(* IEC 61131-3 sources: daoli-st-library/DL_Motion (part 22) *)

(* ---- FB_DL_ElectronicCam.st ---- *)
(*==============================================================================
 * 组件名称 (Component)  : FB_DL_ElectronicCam
 * 所属子库 (Sublibrary) : DL_Motion
 * 当前版本 (Version)    : 1.0.0
 * 组件分类 (Category)   : 功能块（FUNCTION_BLOCK）· 多轴同步耦合族 · 电子凸轮
 * 兼容性   (Platform)   : CODESYS 3.5 / TwinCAT 3 / 汇川 InoProShop / Schneider
 *                         Machine Expert；仅依赖 Standard.library
 *                         （R_TRIG / LIMIT / MIN / MAX / ABS / 类型转换），零厂商方言
 * 接口依赖 (Depends)    : I_DL_MotionAxis / E_DL_AxisState（既有契约，Round 05，零修改）
 * 功能描述 (Function)   : 电子凸轮（PLCopen 凸轮耦合语义的 clean-room 独立实现）。
 *                         以「主轴相位归一化 → 分段线性表插值 → 缩放与偏移」四段
 *                         链计算从轴目标位置，支持周期 / 非周期两种运行方式、主
 *                         轴相位固定偏移与运行相位微调（飞剪切点补偿）、表单调性
 *                         校验与啮合过渡。
 * 设计要点 (Key notes)  :
 *   ① 相位归一化用「截断取整 + 条件加减」实现小数部分，绝不对负数取模，
 *      保证负向主轴时相位仍落在 0.0..1.0。
 *   ② 表查找为线性扫描 + 防死锁计数器；插值斜率计算前强制判分母，重合点保底
 *      取左值（重合已在啮合前由单调性校验拦截）。
 *   ③ 啮合前对全表做一次性扫描（点数 / 单调性 / 非有限值），运行中只校验当前
 *      区间，避免每拍全表扫描拖长任务周期。
 *   ④ 对轴接口每拍至多一次方法调用：定位指令与减速指令在同一拍互斥。
 * 开源溯源 (Origin)     : 原创实现，clean-room。语义来源为汇川 / CODESYS SoftMotion
 *                         公开指令手册的凸轮耦合页面、ABB AC500 PLCopen 库公开
 *                         帮助页、PLC 技术网公开实战帖与非周期追剪技术文
 *                         （来源编号 RAW_NOTES S-2）。
 *                         「借鉴对象的许可说明」：上述对象全部为公开发布但受版权
 *                         保护的帮助文档 / 论坛教程 / 技术文章，属「可免费查阅、
 *                         仅借鉴语义」类别；本实现未复制任何厂商源码、未使用其
 *                         凸轮表 XML 格式，引脚命名、表结构、插值实现、单调性
 *                         校验、故障码与状态机 100% 自有设计。
 * 验收向量 (Acceptance) :
 *   V1 三点表（0/0、180/90、360/0）周期运行：从轴位置连续，无阶跃跳变；
 *   V2 非周期走完表尾 → eComplete 且 bEndOfProfile 置位，等新啮合沿重启；
 *   V3 主轴点等值（非单调）→ 啮合沿受理时锁存 0004_0261；
 *   V4 nCamPoints = 1 → 锁存 0004_0260；
 *   V5 反向主轴 + bDirNegative = TRUE 正常同步；bDirNegative = FALSE 时停留
 *      eWaiting 并出信息级 0004_0140；
 *   V6 fPhaseShift 步进 5 mm → 切点前移且出信息级 0004_0142；
 *   V7 缩放填 0 → 回默认 1.0 并出信息级 0004_0141；
 *   V8 表值含非有限值 → 锁存 0004_0263；
 *   V9 运行中途插入跟踪脉冲 bTrack：重采样相位基准、退回 eIdle（公约 0.1）。
 * 已知限制 (Limits)     :
 *   ① 从轴定位经轴接口每拍一次下发，同步精度受扫描周期限制，属「逻辑层同步」
 *      而非硬实时插补；高速飞剪必须由驱动侧凸轮功能或实时总线插补承载。
 *   ② 不实现分离式凸轮表句柄（表以数组直传，避免句柄生命周期管理）；
 *      不实现凸轮开关量输出（HMI 层量，非运动语义）。
 *   ③ 表数组维度以字面量 16 声明：FB 内部常量不能用于其自身引脚声明，
 *      因此运行期以 UPPER_BOUND 实测维度做二次钳位，实际可用点数不超实测维度。
 *   ④ 相位微调的加减速平滑由调用方斜坡化：本块只检测突变并提示，不代为滤波。
 *   ⑤ 本块为逻辑层同步编排，不构成 ISO 13849 / IEC 62061 认证安全功能。
 * 规格偏离 (Deviation)  :
 *   ① 依公约 0.1 增补 bTrack 输入引脚（首扫 / 跟踪范式强制项）。
 *   ② 表数组声明维度取字面量 16（等同 DL_CAM_MAX_POINTS），理由见已知限制③；
 *      运行期以 UPPER_BOUND / LOWER_BOUND 实测边界做钳位与越界防护。
 *   ③ eDisengaging 每拍重发一次零速指令（受控降速），而非整段只发一次：部分
 *      实现中单次速度指令会被后续局部指令覆盖，逐拍重发更稳妥，且仍满足
 *      「每拍至多一次方法调用」的接口配额。
 *   ④ bEnable 撤除时除清零输出外补发一次停止请求（安全保守处置）。
 *   ⑤ 方向判定对静止主轴（速度绝对值小于判零容差）放行，避免旋转刀从静止
 *      起步时永久停在等待态。
 * 红线自检 (Redline)    :
 *   R1 零全局符号区访问 ✓（无全局变量表访问、无外部变量声明）
 *   R2 零物理地址直写 ✓（无输入输出通道地址记号）
 *   R3 纯 IEC 61131-3 ✓（仅 R_TRIG / LIMIT / MIN / MAX / ABS / 标准类型转换）
 *   R4 防除零 / 防越界 / 浮点容差 ✓（插值前判斜率分母、数组索引经上下界实测
 *      钳位、浮点比较全用 ABS 容差、扫描循环带防死锁计数器）
 *   R5 声明行 100% 中英双语同行注释 ✓
 *   R6 ENUM + CASE 且 CASE 含 ELSE 兜底 ✓
 *   R7 边沿实例无条件周期刷新 ✓（本块无单拍脉冲输出，无跨周期残留标志）
 *   POU 终结符成对 ✓（FUNCTION_BLOCK ↔ END_FUNCTION_BLOCK，末行即终结符；
 *   TYPE ↔ END_TYPE 成对）
 * 故障码表 (Error codes):
 *   16#0004_0140【信息级】主轴方向不符 / 非周期未进表首区，等待中；
 *   16#0004_0141【信息级】缩放系数非法回默认；
 *   16#0004_0142【信息级】相位微调突变超限提示；
 *   16#0004_0260【故障级】凸轮点数非法，锁存；
 *   16#0004_0261【故障级】凸轮表主轴点非单调递增，锁存；
 *   16#0004_0262【故障级】周期长度非法（周期模式），锁存；
 *   16#0004_0263【故障级】凸轮表含非有限值，锁存；
 *   16#0004_0264【故障级】从轴定位指令被拒，锁存；
 *   16#0004_0265【故障级】从轴故障中断耦合（透传），锁存；
 *   16#0004_0298【故障级】非法状态兜底（本块专用，不与其他块共用）。
 *   信息级码只进 uErrorId；bError 为派生式仅反映 eFault 态。
 * 修订历史 (Revision)   :
 *   2026-11-15  v1.0.0  首版入库（Round 08 · DL_Motion 同步耦合族）
 *============================================================================*)

(*-----------------------------------------------------------------------------
 * 调用示例 (Instance guide)：
 *   fbCam.iMaster := fbMasterAxis;                // 主轴实现块实例注入
 *   fbCam.iSlave  := fbSlaveAxis;                 // 从轴实现块实例注入
 *   fbCam.afCamMaster[0] := 0.0;  fbCam.afCamSlave[0] := 0.0;
 *   fbCam.afCamMaster[1] := 180.0; fbCam.afCamSlave[1] := 90.0;
 *   fbCam.afCamMaster[2] := 360.0; fbCam.afCamSlave[2] := 0.0;
 *   fbCam.fCamMasterPeriod := 360.0;
 *   fbCam(bEnable := TRUE, bExecute := bCamCmd, bPeriodic := TRUE,
 *         nCamPoints := 3, fVelLimit := 300.0, fAcc := 2000.0);
 *   注：表数组在周期调用前填好即可（运行中改表无效，须重新啮合）。
 *----------------------------------------------------------------------------*)

(*-----------------------------------------------------------------------------
 * 常见误用与现场提示 (Field notes)：
 *   1 表内主轴点必须严格递增；周期模式下末点可等于周期长度（自然回绕），
 *     但不得小于前一点，否则啮合沿直接被拒（故障级 0261）。
 *   2 相位微调 fPhaseShift 是「运行中」微调量，配方切换请改 fMasterOffset，
 *     两者在块内相加，不会互相覆盖。
 *   3 非周期模式走完表尾后停在 eComplete，必须给新的 bExecute 上升沿才能重启；
 *     周期性连续生产请把 bPeriodic 置 TRUE。
 *   4 等待态与啮合态内本块不会向从轴发停止指令（会与追赶指令打架），要停轴
 *     请给 bDisengage 上升沿，走受控降速路径。
 *   5 主轴静止时相位冻结在最后一次有效值，从轴保持当前位置，属正常工况。
 *----------------------------------------------------------------------------*)

(*-----------------------------------------------------------------------------
 * 枚举: E_DL_CamState（归属 DL_Motion，与本功能块同文件发布）
 * 含义: 电子凸轮耦合状态机，编号间隔 10 预留扩展位。
 *----------------------------------------------------------------------------*)
{attribute 'strict'}
{attribute 'qualified_only'}
TYPE E_DL_CamState :
(
    eIdle        := 0,    // 空闲：未建立耦合，输出指令为零 / Idle: no coupling, command zero
    eWaiting     := 10,   // 等待起步条件：方向不符或未达表首区 / Waiting: direction or table-start condition not met
    eEngaging    := 20,   // 啮合过渡：从轴按速度上限与加速度趋近凸轮目标 / Engaging: slave chases cam target
    eInSync      := 30,   // 同步中：从轴每拍跟随凸轮目标，bInSync 唯一来源 / In sync: slave follows cam target each scan
    eDisengaging := 40,   // 脱开：受控降速后停轴 / Disengaging: controlled deceleration then stop
    eComplete    := 50,   // 非周期走完表尾：bEndOfProfile 有效，等新啮合沿 / Complete: end of profile, waiting for new engage edge
    eFault       := 99    // 故障锁存：仅 bReset 上升沿可退出 / Fault: latched, only bReset rising edge exits
) UINT;
END_TYPE

FUNCTION_BLOCK FB_DL_ElectronicCam
VAR_INPUT
    bEnable         : BOOL := FALSE;        // 总使能（Enable），FALSE=立即脱开并清指令，电平语义
    bExecute        : BOOL := FALSE;        // 建立凸轮耦合（Engage），上升沿受理，仅 eIdle / eComplete 受理
    bDisengage      : BOOL := FALSE;        // 脱开（Disengage），上升沿受理，优先于 bExecute
    bTrack          : BOOL := FALSE;        // 相位基准重同步（Tracking pulse），上升沿即重采样相位基准并退回 eIdle
    bPeriodic       : BOOL := TRUE;         // 周期模式（Periodic），TRUE=表尾回绕表头，FALSE=单程到表尾置完成
    bDirNegative    : BOOL := FALSE;        // 期望主轴方向（Expected master direction），FALSE=正向，TRUE=负向
    fMasterOffset   : REAL := 0.0;          // 主轴相位固定偏移（Master offset）[mm]，配方级参数
    fPhaseShift     : REAL := 0.0;          // 运行相位微调（Phase shift）[mm]，飞剪切点在线补偿，与偏移相加
    fSlaveOffset    : REAL := 0.0;          // 从轴位置偏移（Slave offset）[mm]，叠加在表输出之上
    fMasterScaling  : REAL := 1.0;          // 主轴缩放（Master scaling）[-]，域 0.001..100，非法回默认 1.0
    fSlaveScaling   : REAL := 1.0;          // 从轴缩放（Slave scaling）[-]，域 0.001..100，非法回默认 1.0
    fVelLimit       : REAL := 200.0;        // 从轴速度上限（Slave velocity limit）[mm/s]，域 0.1..100000，兼作定位指令速度
    fAcc            : REAL := 1000.0;       // 从轴加速度（Slave acceleration）[mm/s²]，域 0.1..100000，非有限值回默认
    fDec            : REAL := 1000.0;       // 从轴减速度（Slave deceleration）[mm/s²]，域 0.1..100000，非有限值回默认
    nCamPoints      : UINT := 2;            // 凸轮表有效点数（Active cam points）[-]，域 2..实测表维度，<2 判参数非法
    bReset          : BOOL := FALSE;        // 复位故障（Fault reset），上升沿受理，仅 eFault 态有效
END_VAR
VAR_OUTPUT
    bInSync         : BOOL := FALSE;        // 同步中（In sync），仅 eInSync 态为 TRUE
    bBusy           : BOOL := FALSE;        // 执行中（Busy），等待 / 过渡 / 同步 / 脱开 四态为 TRUE
    bEndOfProfile   : BOOL := FALSE;        // 非周期走完表尾（End of profile），保持到下次啮合受理
    bError          : BOOL := FALSE;        // 故障锁存（Error），派生式仅故障级码参与，信息级码不置位
    uErrorId        : UDINT := 0;           // 故障码（Error code），段位 16#0004_xxxx，0=无故障
    fMasterPhase    : REAL := 0.0;          // 归一化主轴相位（Normalized master phase）[-]，0.0..1.0，HMI 监视用
    fSlavePosCmd    : REAL := 0.0;          // 从轴目标位置指令（Slave position command）[mm]，含缩放与偏移
    fCamSlaveTarget : REAL := 0.0;          // 表插值原始输出（Raw cam output）[mm]，未乘缩放未加偏移，调试用
END_VAR
VAR_IN_OUT
    iMaster         : I_DL_MotionAxis;      // 主轴接口引用（Master axis），由调用方注入实现块实例
    iSlave          : I_DL_MotionAxis;      // 从轴接口引用（Slave axis），由调用方注入实现块实例
    afCamMaster     : ARRAY[0..15] OF REAL; // 凸轮表主轴点（Cam master points）[mm]，维度 16（DL_CAM_MAX_POINTS），须单调递增
    afCamSlave      : ARRAY[0..15] OF REAL; // 凸轮表从轴点（Cam slave points）[mm]，维度 16，与主轴点一一对应
    fCamMasterPeriod: REAL;                 // 周期长度（Master period）[mm]，仅周期模式有效，≤0 判参数非法
END_VAR
VAR
    eState          : E_DL_CamState := E_DL_CamState.eIdle; // 内部状态机步序（Internal state）
    bInit           : BOOL := FALSE;        // 首扫完成标志（First-scan done flag），初值 FALSE，随 bTrack 复位
    bFaultLatch     : BOOL := FALSE;        // 故障锁存标志（Fault latch），仅 bReset 沿或新啮合沿解除
    bTableReady     : BOOL := FALSE;        // 凸轮表就绪标志（Table ready），啮合沿校验通过后置位
    bStopIssued     : BOOL := FALSE;        // 停止请求已发标志（Stop issued flag），单发化防重复发令
    bDirOk          : BOOL := FALSE;        // 主轴方向符合标志（Master direction ok），逐拍重算
    nPtsEff         : DINT := 2;            // 生效点数（Effective point count）[-]，已按实测维度钳位
    nLb             : DINT := 0;            // 表数组下标下界（Array lower bound）[-]，实测取得
    nUb             : DINT := 15;           // 表数组下标上界（Array upper bound）[-]，实测取得
    nAvail          : DINT := 16;           // 实测可用点数（Available points）[-]，上界减下界加一
    iIdx            : DINT := 0;            // 插值区间左端点下标（Interval left index）[-]，已验界
    nIdx            : DINT := 0;            // 表扫描索引（Table scan index）[-]，循环内递增
    nGuard          : DINT := 0;            // 循环防死锁计数器（Loop guard counter）[-]，超限即退出
    fMasterPosEff   : REAL := 0.0;          // 生效主轴坐标（Effective master coordinate）[mm]，含缩放与相位量
    fPhaseRaw       : REAL := 0.0;          // 归一化相位原值（Raw normalized phase）[-]，可为负，需修正
    fPhase          : REAL := 0.0;          // 归一化主轴相位（Normalized phase）[-]，钳在 0.0..1.0
    fPhaseShiftPrev : REAL := 0.0;          // 上拍相位微调量（Previous phase shift）[mm]，突变检测基准
    fKey            : REAL := 0.0;          // 表内主轴求值键（Master key in table）[mm]，已钳到表域
    fM0             : REAL := 0.0;          // 插值区间左主轴点（Interval master low）[mm]
    fM1             : REAL := 0.0;          // 插值区间右主轴点（Interval master high）[mm]
    fS0             : REAL := 0.0;          // 插值区间左从轴点（Interval slave low）[mm]
    fS1             : REAL := 0.0;          // 插值区间右从轴点（Interval slave high）[mm]
    fDen            : REAL := 0.0;          // 插值斜率分母（Interpolation denominator）[mm]，除零前判
    fSlaveTarget    : REAL := 0.0;          // 从轴目标位置（Slave target position）[mm]，含缩放与偏移
    fCamRaw         : REAL := 0.0;          // 表插值原始输出（Raw cam output）[mm]，未加缩放偏移
    fMScaleEff      : REAL := 1.0;          // 生效主轴缩放（Effective master scaling）[-]，非法回 1.0
    fSScaleEff      : REAL := 1.0;          // 生效从轴缩放（Effective slave scaling）[-]，非法回 1.0
    fVelEff         : REAL := 200.0;        // 生效定位速度（Effective velocity）[mm/s]，已做下限兜底
    fAccEff         : REAL := 1000.0;       // 生效加速度（Effective acceleration）[mm/s²]，已做下限兜底
    fDecEff         : REAL := 1000.0;       // 生效减速度（Effective deceleration）[mm/s²]，已做下限兜底
    fPeriodEff      : REAL := 0.0;          // 生效周期长度（Effective period）[mm]，周期模式必须 > 0
    fPosErrBand     : REAL := 0.0;          // 进入同步的位置带宽（Sync band）[mm]，取啮合带宽常量
    fSlavePosNow    : REAL := 0.0;          // 从轴本拍位置（Slave position this scan）[mm]
    fbTrigExec      : R_TRIG;               // 建立耦合指令上升沿（Engage command rising edge）
    fbTrigDisengage : R_TRIG;               // 脱开指令上升沿（Disengage command rising edge）
    fbTrigReset     : R_TRIG;               // 复位指令上升沿（Reset command rising edge）
END_VAR
VAR CONSTANT
    DL_CAM_MAX_POINTS   : DINT := 16;       // 表最大点数（Max table points）[-]，与引脚声明的字面量维度一致
    DL_CAM_INF_MAX      : REAL := 1.0E30;   // 有限值判定幅值上限（Finite magnitude bound）[无量纲，按比较量量纲同值使用]
    DL_CAM_EPS          : REAL := 1.0E-6;   // 浮点判零容差（Float zero tolerance）[无量纲，按比较量量纲同值使用]
    DL_CAM_PAR_FLOOR    : REAL := 1.0E-3;   // 速度/加速度参数下限（Parameter floor）[mm/s 或 mm/s²]
    DL_CAM_VEL_DEF      : REAL := 200.0;    // 速度默认回退值（Default velocity）[mm/s]
    DL_CAM_ACC_DEF      : REAL := 1000.0;   // 加速度默认回退值（Default acceleration）[mm/s²]
    DL_CAM_DEC_DEF      : REAL := 1000.0;   // 减速度默认回退值（Default deceleration）[mm/s²]
    DL_CAM_SCALE_MIN    : REAL := 1.0E-3;   // 缩放系数下限（Scaling floor）[-]，低于此值回默认
    DL_CAM_SCALE_MAX    : REAL := 100.0;    // 缩放系数上限（Scaling ceiling）[-]，高于此值回默认
    DL_CAM_ENGAGE_BAND  : REAL := 0.05;     // 啮合带宽（Engage band）[mm]，位置差进入带宽即判同步
    DL_CAM_PHASE_JUMP   : REAL := 2.0;      // 相位微调突变阈值（Phase jump threshold）[mm]，超此值仅提示
    DL_CAM_END_BAND     : REAL := 0.05;     // 表尾判定带（End band）[mm]，主轴接近末点即判走完
    DL_CAM_GUARD_LIMIT  : DINT := 64;       // 表扫描防死锁上限（Loop guard limit）[-]，远超最大点数
END_VAR

// 段 1｜边沿实例无条件周期刷新（红线 R7：严禁置于 IF / CASE 分支内）
fbTrigExec(CLK := bExecute);
fbTrigDisengage(CLK := bDisengage);
fbTrigReset(CLK := bReset);

// 段 2｜出口默认赋值（公约 0.9：早退路径输出必须确定）
bInSync      := FALSE;
bBusy        := FALSE;
bError       := (eState = E_DL_CamState.eFault);
fSlavePosCmd := 0.0;

// 段 3｜接口引用有效性防御：任一引用未注入则清输出退出，不产生误动作
IF (iMaster = 0) OR (iSlave = 0) THEN
    RETURN;
END_IF

// 段 4｜缩放与速度参数防御（非有限值 / 越域一律回默认并提示，逐拍重算）
IF (fMasterScaling <> fMasterScaling) OR (ABS(fMasterScaling) > DL_CAM_INF_MAX)
   OR (fMasterScaling < DL_CAM_SCALE_MIN) OR (fMasterScaling > DL_CAM_SCALE_MAX) THEN
    fMScaleEff := 1.0;                                   // 主轴缩放非法 → 默认 1.0
    uErrorId   := 16#0004_0141;                          // 【信息级】缩放系数非法回默认
ELSE
    fMScaleEff := fMasterScaling;
END_IF

IF (fSlaveScaling <> fSlaveScaling) OR (ABS(fSlaveScaling) > DL_CAM_INF_MAX)
   OR (fSlaveScaling < DL_CAM_SCALE_MIN) OR (fSlaveScaling > DL_CAM_SCALE_MAX) THEN
    fSScaleEff := 1.0;                                   // 从轴缩放非法 → 默认 1.0
    uErrorId   := 16#0004_0141;                          // 【信息级】缩放系数非法回默认
ELSE
    fSScaleEff := fSlaveScaling;
END_IF

IF (fVelLimit <> fVelLimit) OR (ABS(fVelLimit) > DL_CAM_INF_MAX) OR (fVelLimit < DL_CAM_PAR_FLOOR) THEN
    fVelEff := DL_CAM_VEL_DEF;                           // 速度上限非法 → 默认值
ELSE
    fVelEff := fVelLimit;
END_IF

IF (fAcc <> fAcc) OR (ABS(fAcc) > DL_CAM_INF_MAX) OR (fAcc < DL_CAM_PAR_FLOOR) THEN
    fAccEff := DL_CAM_ACC_DEF;
ELSE
    fAccEff := fAcc;
END_IF

IF (fDec <> fDec) OR (ABS(fDec) > DL_CAM_INF_MAX) OR (fDec < DL_CAM_PAR_FLOOR) THEN
    fDecEff := DL_CAM_DEC_DEF;
ELSE
    fDecEff := fDec;
END_IF

// 段 5｜数组实测边界（公约 0.14：数组访问前必须验界，禁越界索引）
nLb    := LOWER_BOUND(afCamMaster, 1);
nUb    := UPPER_BOUND(afCamMaster, 1);
nAvail := nUb - nLb + 1;
IF nAvail > DL_CAM_MAX_POINTS THEN
    nAvail := DL_CAM_MAX_POINTS;                         // 实测维度超库级上限时按上限钳位，防下标越界
END_IF
IF nAvail < 2 THEN
    nAvail := 0;                                         // 表维度异常（不足两点）时置 0，后续一律判故障
END_IF

// 段 6｜周期长度防御（仅周期模式需要）
IF (fCamMasterPeriod <> fCamMasterPeriod) OR (ABS(fCamMasterPeriod) > DL_CAM_INF_MAX) THEN
    fPeriodEff := 0.0;
ELSE
    fPeriodEff := fCamMasterPeriod;
END_IF

// 段 7｜主轴相位归一化（截断取整 + 条件加减，绝不对负数取模）
fMasterPosEff := fMScaleEff * iMaster.fPosition + fMasterOffset + fPhaseShift;
fPhase        := 0.0;
IF bPeriodic THEN
    IF fPeriodEff > DL_CAM_EPS THEN
        fPhaseRaw := fMasterPosEff / fPeriodEff;         // 分母已验非零
        fPhase    := fPhaseRaw - DINT_TO_REAL(REAL_TO_DINT(fPhaseRaw)); // 截断取整求小数部分
        IF fPhase < 0.0 THEN
            fPhase := fPhase + 1.0;                      // 负向主轴修正到 0.0..1.0
        END_IF
        IF fPhase >= 1.0 THEN
            fPhase := 0.0;                               // 极接近 1.0 的浮点残差归位，防越界
        END_IF
    END_IF
ELSE
    fPhase := 0.0;                                       // 非周期模式不使用归一化相位
END_IF
fMasterPhase := fPhase;

// 段 8｜相位微调突变检测（信息级提示，不阻断；平滑由调用方斜坡化）
IF ABS(fPhaseShift - fPhaseShiftPrev) > DL_CAM_PHASE_JUMP THEN
    uErrorId := 16#0004_0142;                            // 【信息级】相位微调突变超限提示
END_IF
fPhaseShiftPrev := fPhaseShift;

// 段 9｜凸轮表求值（表就绪时逐拍求值；区间右端点下标已由点数钳位保证不越界）
fCamRaw := 0.0;
IF bTableReady AND (nPtsEff >= 2) AND (nPtsEff <= nAvail) THEN
    IF bPeriodic THEN
        // 周期模式：相位展宽到表主轴域（区间端点取实测下标，避免点数与维度不一致）
        fKey := fPhase * (afCamMaster[nLb + nPtsEff - 1] - afCamMaster[nLb]) + afCamMaster[nLb];
    ELSE
        // 非周期模式：主轴坐标钳到表域
        fKey := LIMIT(afCamMaster[nLb], fMasterPosEff, afCamMaster[nLb + nPtsEff - 1]);
    END_IF
    iIdx   := nLb;
    nGuard := 0;
    FOR nIdx := nLb TO (nLb + nPtsEff - 2) DO
        IF nGuard >= DL_CAM_GUARD_LIMIT THEN
            EXIT;                                        // 防死锁：超限退出，保留下标不越界
        END_IF
        nGuard := nGuard + 1;
        iIdx   := nIdx;
        IF fKey <= afCamMaster[nIdx + 1] THEN
            EXIT;                                        // 找到所在区间
        END_IF
    END_FOR
    fM0  := afCamMaster[iIdx];
    fM1  := afCamMaster[iIdx + 1];
    fS0  := afCamSlave[iIdx];
    fS1  := afCamSlave[iIdx + 1];
    fDen := fM1 - fM0;
    IF ABS(fDen) > DL_CAM_EPS THEN
        fCamRaw := fS0 + (fKey - fM0) * (fS1 - fS0) / fDen; // 分段线性插值，分母已验非零
    ELSE
        fCamRaw := fS0;                                  // 区间退化保底取左值（啮合前已被单调性校验拦截）
    END_IF
END_IF
fCamSlaveTarget := fCamRaw;
fSlaveTarget    := fSScaleEff * fCamRaw + fSlaveOffset;

// 段 10｜首扫与跟踪范式（公约 0.1：bTrack OR (NOT bInit) 为唯一判据，禁止反序）
IF bTrack OR (NOT bInit) THEN
    fPhaseShiftPrev := fPhaseShift;                      // 相位微调基准重采样，防跟踪后误报突变
    bTableReady     := FALSE;                            // 表就绪标志复位，须重新啮合校验
    bStopIssued     := FALSE;
    fSlavePosCmd    := 0.0;
    eState          := E_DL_CamState.eIdle;
    bInit           := TRUE;                             // 首扫完成后置位（判据恒为 bTrack OR NOT bInit）
END_IF

// 段 11｜总使能撤除：清零输出并向从轴补发一次停止请求（安全保守处置）
IF NOT bEnable THEN
    IF (NOT bStopIssued) AND ((eState = E_DL_CamState.eEngaging) OR (eState = E_DL_CamState.eInSync)) THEN
        iSlave.Stop();                                   // 使能撤除瞬间单发停止，杜绝残余定位指令
        bStopIssued := TRUE;
    END_IF
    eState       := E_DL_CamState.eIdle;
    bTableReady  := FALSE;
    fSlavePosCmd := 0.0;
END_IF

// 段 12｜事件码管理（公约 0.7 / R15）：锁存码仅在解除路径清，瞬时码逐拍重算
IF NOT bFaultLatch THEN
    uErrorId := 0;
END_IF

// 段 13｜主状态机（ENUM + CASE + ELSE 兜底）
CASE eState OF

    E_DL_CamState.eIdle:                                 // 空闲：等待啮合沿与全表校验
        bBusy := FALSE;
        IF fbTrigExec.Q AND bEnable THEN
            bFaultLatch := FALSE;                        // 新啮合沿：锁存码解除路径（R15）
            bEndOfProfile := FALSE;
            IF (UINT_TO_DINT(nCamPoints) < 2) OR (UINT_TO_DINT(nCamPoints) > nAvail)
               OR (nAvail < 2) THEN
                bFaultLatch := TRUE;
                uErrorId    := 16#0004_0260;             // 【故障级】凸轮点数非法
                eState      := E_DL_CamState.eFault;
            ELSIF bPeriodic AND (fPeriodEff <= DL_CAM_EPS) THEN
                bFaultLatch := TRUE;
                uErrorId    := 16#0004_0262;             // 【故障级】周期长度非法（周期模式）
                eState      := E_DL_CamState.eFault;
            ELSE
                nPtsEff := UINT_TO_DINT(nCamPoints);
                // 啮合前全表一次性扫描：非有限值与单调性（运行中只校验当前区间）
                bTableReady := TRUE;
                nGuard      := 0;
                FOR nIdx := nLb TO (nLb + nPtsEff - 1) DO
                    IF nGuard >= DL_CAM_GUARD_LIMIT THEN
                        EXIT;                            // 防死锁
                    END_IF
                    nGuard := nGuard + 1;
                    IF (afCamMaster[nIdx] <> afCamMaster[nIdx]) OR (afCamSlave[nIdx] <> afCamSlave[nIdx]) THEN
                        bTableReady := FALSE;
                        uErrorId    := 16#0004_0263;     // 【故障级】凸轮表含非有限值
                    END_IF
                END_FOR
                IF bTableReady THEN
                    nGuard := 0;
                    FOR nIdx := nLb TO (nLb + nPtsEff - 2) DO
                        IF nGuard >= DL_CAM_GUARD_LIMIT THEN
                            EXIT;                        // 防死锁
                        END_IF
                        nGuard := nGuard + 1;
                        IF (afCamMaster[nIdx + 1] - afCamMaster[nIdx]) <= DL_CAM_EPS THEN
                            bTableReady := FALSE;
                            uErrorId    := 16#0004_0261; // 【故障级】凸轮表主轴点非单调递增
                        END_IF
                    END_FOR
                END_IF
                IF NOT bTableReady THEN
                    bFaultLatch := TRUE;
                    eState      := E_DL_CamState.eFault;
                ELSE
                    eState := E_DL_CamState.eWaiting;    // 校验通过 → 等待起步条件
                END_IF
            END_IF
        END_IF

    E_DL_CamState.eWaiting:                              // 等待起步条件：方向与表首区
        bBusy := TRUE;
        IF fbTrigDisengage.Q THEN
            eState := E_DL_CamState.eDisengaging;        // 脱开沿优先（本态禁发停止指令）
        ELSIF iSlave.bError THEN
            bFaultLatch := TRUE;
            uErrorId    := 16#0004_0265;                 // 【故障级】从轴故障中断耦合
            eState      := E_DL_CamState.eFault;
        ELSE
            // 方向判定：静止主轴放行（避免旋转刀从静止起步时永久等待）
            IF ABS(iMaster.fVelocity) <= DL_CAM_EPS THEN
                bDirOk := TRUE;
            ELSIF bDirNegative THEN
                bDirOk := (iMaster.fVelocity < 0.0);
            ELSE
                bDirOk := (iMaster.fVelocity > 0.0);
            END_IF
            IF (NOT bDirOk)
               OR ((NOT bPeriodic) AND (fMasterPosEff < afCamMaster[nLb] - DL_CAM_END_BAND)) THEN
                uErrorId := 16#0004_0140;                // 【信息级】方向不符 / 未进表首区，等待中
            ELSE
                eState := E_DL_CamState.eEngaging;
            END_IF
        END_IF

    E_DL_CamState.eEngaging:                             // 啮合过渡：追赶凸轮目标，带宽内转同步
        bBusy := TRUE;
        IF fbTrigDisengage.Q THEN
            eState := E_DL_CamState.eDisengaging;
        ELSIF iSlave.bError THEN
            bFaultLatch := TRUE;
            uErrorId    := 16#0004_0265;                 // 【故障级】从轴故障中断耦合
            eState      := E_DL_CamState.eFault;
        ELSE
            fSlavePosNow := iSlave.fPosition;
            fPosErrBand  := DL_CAM_ENGAGE_BAND;
            IF ABS(fSlavePosNow - fSlaveTarget) <= fPosErrBand THEN
                eState := E_DL_CamState.eInSync;         // 进入带宽 → 同步
            ELSE
                fSlavePosCmd := fSlaveTarget;
                IF NOT iSlave.MoveAbsolute(fPos := fSlaveTarget, fVel := fVelEff, fAcc := fAccEff) THEN
                    bFaultLatch := TRUE;
                    uErrorId    := 16#0004_0264;         // 【故障级】从轴定位指令被拒
                    eState      := E_DL_CamState.eFault;
                END_IF
            END_IF
        END_IF

    E_DL_CamState.eInSync:                               // 同步中：逐拍跟随凸轮目标
        bBusy   := TRUE;
        bInSync := TRUE;
        IF fbTrigDisengage.Q THEN
            eState := E_DL_CamState.eDisengaging;
        ELSIF iSlave.bError THEN
            bFaultLatch := TRUE;
            uErrorId    := 16#0004_0265;                 // 【故障级】从轴故障中断耦合
            eState      := E_DL_CamState.eFault;
        ELSE
            fSlavePosCmd := fSlaveTarget;
            IF NOT iSlave.MoveAbsolute(fPos := fSlaveTarget, fVel := fVelEff, fAcc := fAccEff) THEN
                bFaultLatch := TRUE;
                uErrorId    := 16#0004_0264;             // 【故障级】从轴定位指令被拒
                eState      := E_DL_CamState.eFault;
            ELSIF (NOT bPeriodic) AND (fMasterPosEff >= (afCamMaster[nLb + nPtsEff - 1] - DL_CAM_END_BAND)) THEN
                bEndOfProfile := TRUE;                   // 非周期走完表尾
                bStopIssued   := FALSE;
                eState        := E_DL_CamState.eComplete;
            END_IF
        END_IF

    E_DL_CamState.eDisengaging:                          // 脱开：受控降速后停轴
        bBusy := TRUE;
        IF iSlave.bError THEN
            bFaultLatch := TRUE;
            uErrorId    := 16#0004_0265;                 // 【故障级】从轴故障中断耦合
            eState      := E_DL_CamState.eFault;
        ELSIF ABS(iSlave.fVelocity) <= DL_CAM_EPS THEN
            IF NOT bStopIssued THEN
                iSlave.Stop();                           // 已停稳：单发停止确认（本拍唯一一次轴调用）
                bStopIssued := TRUE;
            END_IF
            fSlavePosCmd := 0.0;
            bBusy        := FALSE;
            bStopIssued  := FALSE;                       // 停发标志闭环复位
            eState       := E_DL_CamState.eIdle;
        ELSE
            // 逐拍重发零速指令保证持续减速（每拍至多一次轴调用）
            IF NOT iSlave.MoveVelocity(fVel := 0.0, fAcc := fDecEff) THEN
                bFaultLatch := TRUE;
                uErrorId    := 16#0004_0264;             // 【故障级】脱开减速指令被拒
                eState      := E_DL_CamState.eFault;
            END_IF
            fSlavePosCmd := 0.0;
        END_IF

    E_DL_CamState.eComplete:                             // 非周期完成：保持结果等新啮合沿
        bBusy         := FALSE;
        bEndOfProfile := TRUE;
        fSlavePosCmd  := fSlaveTarget;                   // 保持末点目标，从轴稳定停在表尾位置
        IF fbTrigDisengage.Q THEN
            eState := E_DL_CamState.eDisengaging;
        ELSIF fbTrigExec.Q AND bEnable THEN
            bEndOfProfile := FALSE;                      // 新啮合沿受理：清完成标志重新起步
            bFaultLatch   := FALSE;
            eState        := E_DL_CamState.eWaiting;
        END_IF

    E_DL_CamState.eFault:                                // 故障锁存：仅复位沿可退出
        bBusy         := FALSE;
        bInSync       := FALSE;
        fSlavePosCmd  := 0.0;
        bStopIssued   := FALSE;
        bTableReady   := FALSE;
        IF fbTrigReset.Q THEN
            bFaultLatch := FALSE;                        // 唯一解除路径
            uErrorId    := 0;
            bEndOfProfile := FALSE;
            eState      := E_DL_CamState.eIdle;
        END_IF

    ELSE                                                 // 非法状态兜底（本块专用码）
        bFaultLatch   := TRUE;
        uErrorId      := 16#0004_0298;                   // 【故障级】非法状态兜底
        bBusy         := FALSE;
        bInSync       := FALSE;
        bTableReady   := FALSE;
        fSlavePosCmd  := 0.0;
        eState        := E_DL_CamState.eFault;

END_CASE

// 段 14｜出口映射（派生式，信息级码不参与 bError）
bError          := (eState = E_DL_CamState.eFault);
bInSync         := (eState = E_DL_CamState.eInSync);
bBusy           := (eState = E_DL_CamState.eWaiting) OR (eState = E_DL_CamState.eEngaging)
                   OR (eState = E_DL_CamState.eInSync) OR (eState = E_DL_CamState.eDisengaging);
fCamSlaveTarget := fCamRaw;
fMasterPhase    := fPhase;

END_FUNCTION_BLOCK

(* ---- FB_DL_ElectronicGear.st ---- *)
(*==============================================================================
 * 组件名称 (Component)  : FB_DL_ElectronicGear
 * 所属子库 (Sublibrary) : DL_Motion
 * 当前版本 (Version)    : 1.0.0
 * 组件分类 (Category)   : 功能块（FUNCTION_BLOCK）· 多轴同步耦合族 · 电子齿轮
 * 兼容性   (Platform)   : CODESYS 3.5 / TwinCAT 3 / 汇川 InoProShop / Schneider
 *                         Machine Expert；仅依赖 Standard.library
 *                         （R_TRIG / LIMIT / MIN / MAX / ABS），零厂商方言
 * 接口依赖 (Depends)    : I_DL_MotionAxis / E_DL_AxisState（既有契约，Round 05，
 *                         零修改引用；本块不新增任何接口方法）
 * 功能描述 (Function)   : 电子齿轮耦合（PLCopen 齿轮耦合语义的 clean-room 独立
 *                         实现）。从轴速度指令 = 主轴实际速度 × 传动比 + 相位
 *                         补偿项。传动比以整数分子/分母保存，仅在输出处换算为
 *                         浮点比值，避免浮点比值累积误差；啮合过渡段按 fAcc 限
 *                         斜率平滑建立，脱开段按 fDec 受控降速到零后再向轴发一次
 *                         停止请求。
 * 设计要点 (Key notes)  :
 *   ① 整数比值对：nRatioNum / nRatioDen 全程整数保存，fRatio 仅为显示量；
 *      分数比 3:7 长期运行不产生浮点漂移（验收向量 V2）。
 *   ② 相位补偿为比例式（fPhaseGain × 累计相位误差，钳到 ±fPhaseMax），
 *      不在轴外层再套积分器；fPhaseGain = 0 时补偿恒为 0（功能关闭）。
 *   ③ 指令下发去抖：仅当新指令与上次下发值之差超过重发阈值才向从轴下发，
 *      避免每拍刷指令洪水（接口配额：对轴接口每拍至多一次方法调用）。
 *   ④ 连续更新门控：eInGear 内改传动比，未开放连续更新时拒绝并出信息级码。
 * 开源溯源 (Origin)     : 原创实现，clean-room。语义来源为 PLCopen
 *                         「Function blocks for motion control」公开规范
 *                         （MC_GearIn / MC_GearInPos 引脚表与状态语义）、
 *                         infoPLC 公开镜像的 Part 2 扩展版说明、Beckhoff
 *                         TF5200 编程手册公开帮助页、Unitronics 多轴指令公开
 *                         帮助页（来源编号 RAW_NOTES S-1）。
 *                         「借鉴对象的许可说明」：上述对象均为公开发布但受版权
 *                         保护的规范文档 / 厂商帮助文档，属「可免费查阅、
 *                         可借鉴接口参数域与状态语义、禁止复制代码」类别；本
 *                         实现未复制任何示例代码、源码行或表结构，引脚命名、
 *                         枚举、状态机跃迁、故障码、相位补偿控制律 100% 自有。
 * 验收向量 (Acceptance) :
 *   V1 正常啮合：比值 1:2、主速 100 → 从速指令趋近 200，过渡段每拍增速不超
 *      fAcc × 采样周期；
 *   V2 分数比 3:7 长期运行：fRatio 恒为 0.428571（整数比值不漂移），相位误差
 *      有界不发散；
 *   V3 分母 0：bExecute 沿受理时判参数非法 → 锁存 0004_0250，指令清零不进耦合；
 *   V4 bContinuousUpdate = FALSE 时改比值：沿用旧比值 + 信息级 0004_0131；
 *   V5 相位补偿开（fPhaseGain = 2）注入 1 mm 相位差：补偿量不超 fPhaseMax，
 *      相位误差单调收敛；
 *   V6 脱开：bDisengage 沿 → 受控降速，指令归零后向轴发一次停止请求 → eIdle；
 *   V7 从轴故障：iSlave.bError 置位 → 锁存 0004_0252 并清指令；
 *   V8 主轴静止：主速绝对值小于判零容差 → 相位积累冻结 + 信息级 0004_0130，
 *      不置故障；
 *   V9 运行中途插入跟踪脉冲 bTrack：重采样主从参考位置、相位误差清零、
 *      耦合状态退回 eIdle（公约 0.1 必测向量）。
 * 已知限制 (Limits)     :
 *   ① 主轴与从轴若被注入同一实例，本块无法在块内识别（接口引用不可比较
 *      身份），轴自身仲裁；调用方必须保证主从不指向同一实例。
 *   ② 本库接口无「指令速度」属性，耦合一律取主轴实际速度（等效于按实际值
 *      耦合）；指令值耦合留待接口升版，避免破坏既有 6 个实现块。
 *   ③ 本块为逻辑层同步编排，不构成 ISO 13849 / IEC 62061 认证安全功能；
 *      安全回路、硬限位与机械保护由认证安全控制器与硬件承载。
 *   ④ 同步精度受扫描周期限制，属逻辑层耦合而非硬实时插补。
 * 规格偏离 (Deviation)  :
 *   ① 依公约 0.1（首扫范式）增补 bTrack 输入引脚；依公约 0.10（定时基准由
 *      引脚给）增补 tCycle 输入引脚。二者均为公共约定强制项，非逐组件条款
 *      可覆盖。影响：调用方须接扫描周期常量与跟踪脉冲，其余引脚语义不变。
 *   ② 出口默认赋值置于参数防御之前（依公约 0.9「早退路径输出确定」），与
 *      规格 1.1 节「防御 → 默认」的叙述顺序有调整，语义等价。
 *   ③ bEnable 撤除时除清零输出外，另向从轴补发一次停止请求（安全保守处置：
 *      仅清指令会让从轴保留末次速度指令，现场不可接受）。
 *   ④ 啮合完成判据取「指令与目标之差进入啮合判定带」这一明确口径（带值 0.01 mm/s），
 *      规格原文写「差小于速度上限或绝对值超差小于判零容差十倍」，两种表述在
 *      限速非零时不等价；本实现取固定小带，语义更严（只在真正跟上时才判啮合）。
 * 红线自检 (Redline)    :
 *   R1 零全局符号区访问 ✓（无全局变量表访问、无外部变量声明）
 *   R2 零物理地址直写 ✓（无输入输出通道地址记号）
 *   R3 纯 IEC 61131-3 ✓（仅标准库 R_TRIG / LIMIT / MIN / MAX / ABS / 类型转换）
 *   R4 防除零 / 防越界 / 浮点容差 ✓（比值换算前判分母、浮点比较全用 ABS 容差）
 *   R5 声明行 100% 中英双语同行注释 ✓
 *   R6 ENUM + CASE 且 CASE 含 ELSE 兜底 ✓
 *   R7 边沿实例无条件周期刷新 ✓（R25 单拍闭环：本块无单拍脉冲输出）
 *   POU 终结符成对 ✓（FUNCTION_BLOCK ↔ END_FUNCTION_BLOCK，末行即终结符；
 *   TYPE ↔ END_TYPE 成对）
 * 故障码表 (Error codes):
 *   16#0004_0130【信息级】主轴静止、相位跟踪冻结，不置故障位；
 *   16#0004_0131【信息级】未开放连续更新时改传动比被拒，沿用旧比值；
 *   16#0004_0132【信息级】从轴速度指令被绝对限速钳位；
 *   16#0004_0250【故障级】传动比参数非法（分母为 0 / 分子非正），锁存；
 *   16#0004_0251【故障级】从轴速度指令被轴拒绝，锁存；
 *   16#0004_0252【故障级】从轴故障中断耦合（透传），锁存；
 *   16#0004_0299【故障级】非法状态兜底（本块专用，不与其他块共用）。
 *   信息级码只进 uErrorId，不参与 bError 派生；bError 仅反映 eFault 态。
 * 修订历史 (Revision)   :
 *   2026-11-15  v1.0.0  首版入库（Round 08 · DL_Motion 同步耦合族开族件）
 *============================================================================*)

(*-----------------------------------------------------------------------------
 * 调用示例 (Instance guide)：
 *   fbGear.iMaster := fbMasterAxis;              // 主轴实现块实例注入
 *   fbGear.iSlave  := fbSlaveAxis;               // 从轴实现块实例注入
 *   fbGear(bEnable := TRUE, bExecute := bCoupleCmd,   // 周期调用，永远每拍调用
 *          nRatioNum := 1, nRatioDen := 2,
 *          fAcc := 800.0, fDec := 800.0,
 *          fVelLimit := 600.0, fPhaseGain := 1.5,
 *          tCycle := T#10MS);
 *   IF fbGear.bInGear THEN bReady := TRUE; END_IF
 *   注：从轴速度指令经 fSlaveSpeedCmd 出口逐拍刷新，实际下发由本块内部完成
 *       （每拍至多一次速度指令），上层不要再对同一从轴另发运动指令。
 *----------------------------------------------------------------------------*)

(*-----------------------------------------------------------------------------
 * 常见误用与现场提示 (Field notes)：
 *   1 本块是「速度耦合」而非「位置同步」：位置偏差靠相位补偿项收敛，若现场
 *     需要硬位置对齐（GearInPos 语义），请改用电子凸轮块承载。
 *   2 比值引脚为整数：若工艺给的是小数比值（如 0.28），请放大为整数对
 *     （28 : 100），不要直接填浮点近似值，否则长期运行会漂。
 *   3 主轴静止时相位冻结属正常工况（信息级 0130），不要当作故障处理；
 *     主轴重新启动后相位继续累计。
 *   4 从轴被外部强制停止（驱动器使能丢失）时会锁存 0252；必须等从轴恢复且
 *     给 bReset 上升沿后才能重新啮合。
 *   5 bTrack 用于调试与换型：给一个上升沿即重采样参考位置并退回 eIdle，
 *     不会向从轴发停止请求，轴保持当前运动状态（由调用方决定是否先停轴）。
 *----------------------------------------------------------------------------*)

(*-----------------------------------------------------------------------------
 * 枚举: E_DL_GearState（归属 DL_Motion，与本功能块同文件发布）
 * 含义: 电子齿轮耦合状态机，编号间隔 10 预留扩展位。
 *----------------------------------------------------------------------------*)
{attribute 'strict'}
{attribute 'qualified_only'}
TYPE E_DL_GearState :
(
    eIdle          := 0,    // 空闲：从轴不受本块控制，速度指令清零 / Idle: slave not controlled, speed command cleared
    eSynchronizing := 10,   // 啮合过渡：从轴速度指令向目标比值速度按加速度斜坡逼近 / Synchronizing: slave speed ramps toward ratio target
    eInGear        := 20,   // 已啮合：主从速度比稳定保持，bInGear 唯一来源 / In gear: ratio held steady, sole source of bInGear
    eDisengaging   := 30,   // 脱开：按脱开减速度受控降速至零 / Disengaging: controlled deceleration to zero
    eFault         := 99    // 故障锁存：仅 bReset 上升沿可退出 / Fault: latched, only bReset rising edge exits
) UINT;
END_TYPE

FUNCTION_BLOCK FB_DL_ElectronicGear
VAR_INPUT
    bEnable           : BOOL := FALSE;          // 耦合总使能（Coupling enable），FALSE=脱开并清零输出，电平语义
    bExecute          : BOOL := FALSE;          // 建立耦合指令（Engage command），上升沿受理，eInGear 期间忽略新沿
    bDisengage        : BOOL := FALSE;          // 脱开指令（Disengage command），上升沿受理，优先于 bExecute
    bTrack            : BOOL := FALSE;          // 参考位置重同步（Tracking pulse），上升沿/电平即重采样主从位置并清相位误差
    nRatioNum         : DINT := 1;              // 传动比分子（Gear ratio numerator）[-]，域 1..1000000，≤0 判参数非法
    nRatioDen         : DINT := 1;              // 传动比分母（Gear ratio denominator）[-]，域 1..1000000，=0 防除零故障
    bContinuousUpdate : BOOL := FALSE;          // 运行中改比值使能（Continuous update），FALSE 时啮合内改比值被拒并出信息码
    fAcc              : REAL := 500.0;          // 啮合过渡加速度（Engage acceleration）[mm/s²]，域 0.1..100000，非有限值→默认
    fDec              : REAL := 500.0;          // 脱开减速度（Disengage deceleration）[mm/s²]，域 0.1..100000，非有限值→默认
    fVelLimit         : REAL := 0.0;            // 从轴速度绝对上限（Slave speed limit）[mm/s]，0=不限，负值取绝对值
    fPhaseGain        : REAL := 0.0;            // 相位修正增益（Phase correction gain）[1/s]，0=关闭相位补偿
    fPhaseMax         : REAL := 5.0;            // 相位修正量上限（Phase correction limit）[mm/s]，仅补偿开启时有效
    tCycle            : TIME := T#10MS;         // 任务扫描周期（Task cycle time）[ms]，由调用方按实际任务给，用于加速度限斜率
    bReset            : BOOL := FALSE;          // 复位故障（Fault reset），上升沿受理，仅 eFault 态有效
END_VAR
VAR_OUTPUT
    bInGear           : BOOL := FALSE;          // 已啮合标志（In gear），仅 eInGear 态为 TRUE
    bBusy             : BOOL := FALSE;          // 执行中（Busy），eSynchronizing / eInGear / eDisengaging 为 TRUE
    bActive           : BOOL := FALSE;          // 本块持有从轴控制权（Active），eSynchronizing / eInGear 为 TRUE
    bError            : BOOL := FALSE;          // 故障锁存（Error），派生式仅故障级码参与，信息级码不置位
    uErrorId          : UDINT := 0;             // 故障码（Error code），段位 16#0004_xxxx，0=无故障
    fRatio            : REAL := 0.0;            // 实际生效传动比（Effective ratio）[-]，= 生效分子 / 生效分母
    fSlaveSpeedCmd    : REAL := 0.0;            // 下发给从轴的速度指令（Slave speed command）[mm/s]，带符号，负值=负向
    fPhaseError       : REAL := 0.0;            // 相位累计误差（Accumulated phase error）[mm]，= 累计(主位增量×比值 − 从位增量)
END_VAR
VAR_IN_OUT
    iMaster           : I_DL_MotionAxis;        // 主轴接口引用（Master axis），由调用方注入实现块实例
    iSlave            : I_DL_MotionAxis;        // 从轴接口引用（Slave axis），由调用方注入实现块实例
END_VAR
VAR
    eState            : E_DL_GearState := E_DL_GearState.eIdle; // 内部状态机步序（Internal state）
    bInit             : BOOL := FALSE;          // 首扫完成标志（First-scan done flag），初值 FALSE，随 bTrack 复位重采样
    bFaultLatch       : BOOL := FALSE;          // 故障锁存标志（Fault latch），仅 bReset 沿或新啮合沿解除
    bRatioOk          : BOOL := FALSE;          // 传动比参数合法标志（Ratio parameter valid），逐拍重算
    bStopIssued       : BOOL := FALSE;          // 脱开停止请求已发标志（Stop issued flag），单发化防重复发令
    nNumEff           : DINT := 1;              // 生效传动比分子（Effective numerator）[-]，啮合时锁定
    nDenEff           : DINT := 1;              // 生效传动比分母（Effective denominator）[-]，啮合时锁定且已验非零
    fRatioEff         : REAL := 1.0;            // 生效传动比数值（Effective ratio value）[-]，仅由整数对比值换算
    fAccEff           : REAL := 500.0;          // 生效啮合加速度（Effective acceleration）[mm/s²]，已做默认回退与限幅
    fDecEff           : REAL := 500.0;          // 生效脱开减速度（Effective deceleration）[mm/s²]，已做默认回退与限幅
    fVelLimitEff      : REAL := 0.0;            // 生效速度上限（Effective speed limit）[mm/s]，0=不限
    fPhaseMaxEff      : REAL := 5.0;            // 生效相位补偿上限（Effective phase limit）[mm/s]，≥0
    fDtS              : REAL := 0.01;           // 采样周期秒值（Cycle time in seconds）[s]，由 tCycle 换算并限幅
    fCmdRamp          : REAL := 0.0;            // 斜坡中的速度指令（Ramped speed command）[mm/s]，带符号
    fLastSentCmd      : REAL := 0.0;            // 上次实际下发速度（Last issued speed）[mm/s]，用于重发去抖
    fTargetCmd        : REAL := 0.0;            // 本拍目标速度（Target speed this scan）[mm/s]，含相位补偿与限幅
    fCompTerm         : REAL := 0.0;            // 相位补偿项（Phase compensation term）[mm/s]，已钳到 ±fPhaseMax
    fStepMax          : REAL := 0.0;            // 单拍速度增量上限（Max speed step per scan）[mm/s]，= 加速度 × 采样周期
    fMasterVel        : REAL := 0.0;            // 主轴实际速度（Master actual velocity）[mm/s]，带符号
    fSlaveVel         : REAL := 0.0;            // 从轴实际速度（Slave actual velocity）[mm/s]，带符号
    fMasterPosNow     : REAL := 0.0;            // 主轴本拍位置（Master position this scan）[mm]
    fSlavePosNow      : REAL := 0.0;            // 从轴本拍位置（Slave position this scan）[mm]
    fLastMasterPos    : REAL := 0.0;            // 上拍主轴位置（Previous master position）[mm]，相位增量基准
    fLastSlavePos     : REAL := 0.0;            // 上拍从轴位置（Previous slave position）[mm]，相位增量基准
    fPhaseErrInt      : REAL := 0.0;            // 相位误差累计器（Phase error accumulator）[mm]，内部量
    fNewRatio         : REAL := 1.0;            // 新比值候选值（Candidate ratio value）[-]，除法前已验分母
    fbTrigExec        : R_TRIG;                 // 建立耦合指令上升沿（Engage command rising edge）
    fbTrigDisengage   : R_TRIG;                 // 脱开指令上升沿（Disengage command rising edge）
    fbTrigReset       : R_TRIG;                 // 复位指令上升沿（Reset command rising edge）
END_VAR
VAR CONSTANT
    DL_GEAR_INF_MAX    : REAL := 1.0E30;        // 有限值判定幅值上限（Finite magnitude bound）[无量纲，按各量量纲同值使用]
    DL_GEAR_EPS        : REAL := 1.0E-6;        // 浮点判零容差（Float zero tolerance）[无量纲，按比较量量纲同值使用]
    DL_GEAR_PAR_FLOOR  : REAL := 1.0E-3;        // 加速度/减速度参数下限（Acceleration floor）[mm/s²]，低于此值回默认
    DL_GEAR_ACC_DEF    : REAL := 500.0;         // 加速度默认回退值（Default acceleration）[mm/s²]
    DL_GEAR_DEC_DEF    : REAL := 500.0;         // 减速度默认回退值（Default deceleration）[mm/s²]
    DL_GEAR_ACC_MAX    : REAL := 100000.0;      // 加速度上限（Acceleration upper bound）[mm/s²]，超限钳位
    DL_GEAR_LOCK_BAND  : REAL := 0.01;          // 啮合判定带（In-gear band）[mm/s]，指令与目标差小于此值判啮合
    DL_GEAR_RESEND_EPS : REAL := 0.5;           // 速度指令重发阈值（Resend threshold）[mm/s]，差小于此值不重复下发
    DL_GEAR_DT_MIN     : REAL := 1.0E-4;        // 采样周期下限（Cycle time lower bound）[s]，低于此值按默认
    DL_GEAR_DT_MAX     : REAL := 1.0;           // 采样周期上限（Cycle time upper bound）[s]，高于此值钳位
    DL_GEAR_DT_DEF     : REAL := 0.01;          // 采样周期默认值（Default cycle time）[s]
    DL_GEAR_RATIO_MAX  : DINT := 1000000;       // 传动比分子分母上限（Ratio term upper bound）[-]
END_VAR

// 段 1｜边沿实例无条件周期刷新（红线 R7：严禁置于 IF / CASE 分支内）
fbTrigExec(CLK := bExecute);
fbTrigDisengage(CLK := bDisengage);
fbTrigReset(CLK := bReset);

// 段 2｜出口默认赋值（公约 0.9：早退路径输出必须确定）
bInGear        := FALSE;
bBusy          := FALSE;
bActive        := FALSE;
bError         := (eState = E_DL_GearState.eFault);
fSlaveSpeedCmd := 0.0;
fRatio         := fRatioEff;

// 段 3｜接口引用有效性防御：任一引用未注入则清输出退出，不产生误动作
IF (iMaster = 0) OR (iSlave = 0) THEN
    RETURN;
END_IF

// 段 4｜采样周期换算与限幅（公约 0.10：定时基准由引脚给，禁读系统时钟）
fDtS := TIME_TO_REAL(tCycle) * 1.0E-3;                       // 毫秒 → 秒（注释：本行换算单位为 s）
IF (fDtS <> fDtS) OR (fDtS <= DL_GEAR_DT_MIN) THEN
    fDtS := DL_GEAR_DT_DEF;                                  // 周期非法回默认 10 ms，防除零与超大单拍步长
ELSIF fDtS > DL_GEAR_DT_MAX THEN
    fDtS := DL_GEAR_DT_MAX;                                  // 周期过大钳位，避免单拍跨越过大
END_IF

// 段 5｜参数防御：非有限值回默认、加速度/减速度非正回默认、限速负值取绝对值
IF (fAcc <> fAcc) OR (ABS(fAcc) > DL_GEAR_INF_MAX) OR (fAcc <= DL_GEAR_PAR_FLOOR) THEN
    fAccEff := DL_GEAR_ACC_DEF;                              // 加速度非法 → 默认值
ELSE
    fAccEff := MIN(fAcc, DL_GEAR_ACC_MAX);                   // 加速度合法 → 上限钳位
END_IF

IF (fDec <> fDec) OR (ABS(fDec) > DL_GEAR_INF_MAX) OR (fDec <= DL_GEAR_PAR_FLOOR) THEN
    fDecEff := DL_GEAR_DEC_DEF;                              // 减速度非法 → 默认值
ELSE
    fDecEff := MIN(fDec, DL_GEAR_ACC_MAX);                   // 减速度合法 → 上限钳位
END_IF

IF (fVelLimit <> fVelLimit) OR (ABS(fVelLimit) > DL_GEAR_INF_MAX) THEN
    fVelLimitEff := 0.0;                                     // 限速非有限值 → 视为不限
ELSE
    fVelLimitEff := ABS(fVelLimit);                          // 限速取绝对值，0=不限
END_IF

IF (fPhaseMax <> fPhaseMax) OR (ABS(fPhaseMax) > DL_GEAR_INF_MAX) THEN
    fPhaseMaxEff := 0.0;                                     // 补偿上限非法 → 关闭补偿
ELSE
    fPhaseMaxEff := ABS(fPhaseMax);                          // 补偿上限取绝对值，0=关闭补偿
END_IF

// 传动比参数合法性：分子必须为正、分母必须为正（分母为 0 防除零，负值无工程意义）
bRatioOk := (nRatioNum > 0) AND (nRatioDen > 0)
            AND (nRatioNum <= DL_GEAR_RATIO_MAX) AND (nRatioDen <= DL_GEAR_RATIO_MAX);

// 段 6｜首扫与跟踪范式（公约 0.1：bTrack OR (NOT bInit) 为唯一判据，禁止反序）
fMasterPosNow := iMaster.fPosition;
fSlavePosNow  := iSlave.fPosition;
fMasterVel    := iMaster.fVelocity;
fSlaveVel     := iSlave.fVelocity;

IF bTrack OR (NOT bInit) THEN
    fLastMasterPos := fMasterPosNow;                         // 主轴参考位置重采样 [mm]
    fLastSlavePos  := fSlavePosNow;                          // 从轴参考位置重采样 [mm]
    fPhaseErrInt   := 0.0;                                   // 相位误差清零 [mm]
    fCmdRamp       := fSlaveVel;                             // 斜坡起点取从轴当前速度，避免指令跳变 [mm/s]
    fLastSentCmd   := fSlaveVel;                             // 下发基准同步，避免首拍误判重发 [mm/s]
    bStopIssued    := FALSE;                                 // 停止单发标志复位
    eState         := E_DL_GearState.eIdle;                  // 跟踪后退回空闲，等待新的啮合沿
    bInit          := TRUE;                                  // 首扫完成后置位（判据恒为 bTrack OR NOT bInit）
END_IF

// 段 7｜总使能撤除：清零输出并向从轴补发一次停止请求（安全保守处置）
IF NOT bEnable THEN
    IF (NOT bStopIssued) AND ((eState = E_DL_GearState.eSynchronizing) OR (eState = E_DL_GearState.eInGear)) THEN
        iSlave.Stop();                                       // 使能撤除瞬间单发一次停止，杜绝残余速度指令
        bStopIssued := TRUE;
    END_IF
    eState       := E_DL_GearState.eIdle;
    fCmdRamp     := 0.0;
    fLastSentCmd := 0.0;
    fPhaseErrInt := 0.0;
    fSlaveSpeedCmd := 0.0;
END_IF

// 段 8｜事件码管理（公约 0.7 / R15）：锁存码仅在解除路径清，瞬时码逐拍重算
IF NOT bFaultLatch THEN
    uErrorId := 0;                                           // 非锁存态每拍重算瞬时码
END_IF

// 段 9｜主状态机（ENUM + CASE + ELSE 兜底）
CASE eState OF

    E_DL_GearState.eIdle:                                    // 空闲：等待啮合沿与参数门禁
        bInGear := FALSE;
        bBusy   := FALSE;
        bActive := FALSE;
        IF fbTrigExec.Q AND bEnable THEN
            bFaultLatch := FALSE;                            // 新啮合沿：锁存码解除路径（R15）
            IF NOT bRatioOk THEN
                bFaultLatch    := TRUE;                      // 传动比非法：故障级锁存
                uErrorId       := 16#0004_0250;              // 【故障级】传动比参数非法
                eState         := E_DL_GearState.eFault;
            ELSE
                nNumEff     := nRatioNum;                    // 锁定分子，运行中不受引脚抖动影响
                nDenEff     := nRatioDen;                    // 锁定分母（已验非零）
                fRatioEff   := DINT_TO_REAL(nNumEff) / DINT_TO_REAL(nDenEff); // 整数对比值换算，唯一除法点且分母已验非零
                fRatio      := fRatioEff;
                fCmdRamp    := fSlaveVel;                    // 过渡斜坡起点 = 从轴当前速度
                fLastSentCmd:= fSlaveVel;
                fPhaseErrInt:= 0.0;                          // 新啮合：相位误差从零起算
                bStopIssued := FALSE;
                eState      := E_DL_GearState.eSynchronizing;
            END_IF
        END_IF

    E_DL_GearState.eSynchronizing:                           // 啮合过渡：按加速度限斜率逼近目标比值速度
        bBusy   := TRUE;
        bActive := TRUE;
        IF fbTrigDisengage.Q THEN
            eState := E_DL_GearState.eDisengaging;           // 脱开沿优先于一切运行逻辑
        ELSIF iSlave.bError THEN
            bFaultLatch := TRUE;                             // 从轴故障透传：故障级锁存
            uErrorId    := 16#0004_0252;                     // 【故障级】从轴故障中断耦合
            fCmdRamp    := 0.0;
            fSlaveSpeedCmd := 0.0;
            eState      := E_DL_GearState.eFault;
        ELSE
            // 相位累计：主轴位移增量 × 比值 − 从轴位移增量（主静止时冻结）
            IF ABS(fMasterVel) > DL_GEAR_EPS THEN
                fPhaseErrInt := fPhaseErrInt + (fMasterPosNow - fLastMasterPos) * fRatioEff
                                - (fSlavePosNow - fLastSlavePos);
            ELSE
                uErrorId := 16#0004_0130;                    // 【信息级】主轴静止、相位跟踪冻结（正常工况）
            END_IF
            // 目标速度 = 主速 × 比值 + 相位补偿项
            fCompTerm := 0.0;
            IF (ABS(fPhaseGain) > DL_GEAR_EPS) AND (fPhaseMaxEff > DL_GEAR_EPS) THEN
                fCompTerm := LIMIT(-fPhaseMaxEff, fPhaseGain * fPhaseErrInt, fPhaseMaxEff); // 补偿量钳到 ±上限
            END_IF
            fTargetCmd := fMasterVel * fRatioEff + fCompTerm;
            // 绝对限速钳位（提示配方比值与限速矛盾，逐拍重算不置故障）
            IF (fVelLimitEff > DL_GEAR_EPS) AND (ABS(fTargetCmd) > fVelLimitEff) THEN
                fTargetCmd := LIMIT(-fVelLimitEff, fTargetCmd, fVelLimitEff);
                uErrorId   := 16#0004_0132;                  // 【信息级】从轴速度指令被限速钳位
            END_IF
            // 加速度限斜率：单拍增量不超 加速度 × 采样周期
            fStepMax  := fAccEff * fDtS;
            fCmdRamp  := fCmdRamp + LIMIT(-fStepMax, fTargetCmd - fCmdRamp, fStepMax);
            fSlaveSpeedCmd := fCmdRamp;
            // 每拍至多一次速度指令下发，且仅在变化超过重发阈值时下发
            IF ABS(fCmdRamp - fLastSentCmd) > DL_GEAR_RESEND_EPS THEN
                IF NOT iSlave.MoveVelocity(fVel := fCmdRamp, fAcc := fAccEff) THEN
                    bFaultLatch := TRUE;                     // 指令被轴拒绝：故障级锁存
                    uErrorId    := 16#0004_0251;             // 【故障级】从轴速度指令被拒
                    fCmdRamp    := 0.0;
                    fSlaveSpeedCmd := 0.0;
                    eState      := E_DL_GearState.eFault;
                ELSE
                    fLastSentCmd := fCmdRamp;
                END_IF
            END_IF
            // 指令进入啮合判定带 → 已啮合
            IF (eState = E_DL_GearState.eSynchronizing) AND (ABS(fCmdRamp - fTargetCmd) <= DL_GEAR_LOCK_BAND) THEN
                eState := E_DL_GearState.eInGear;
            END_IF
        END_IF

    E_DL_GearState.eInGear:                                  // 已啮合：比值稳定保持 + 连续更新门控
        bBusy    := TRUE;
        bActive  := TRUE;
        bInGear  := TRUE;
        IF fbTrigDisengage.Q THEN
            eState := E_DL_GearState.eDisengaging;           // 脱开沿优先
        ELSIF iSlave.bError THEN
            bFaultLatch := TRUE;
            uErrorId    := 16#0004_0252;                     // 【故障级】从轴故障中断耦合
            fCmdRamp    := 0.0;
            fSlaveSpeedCmd := 0.0;
            eState      := E_DL_GearState.eFault;
        ELSE
            // 传动比变更门控：未开放连续更新时拒绝，沿用旧比值并出信息码
            IF (nRatioNum <> nNumEff) OR (nRatioDen <> nDenEff) THEN
                IF bContinuousUpdate THEN
                    IF bRatioOk THEN
                        nNumEff   := nRatioNum;
                        nDenEff   := nRatioDen;
                        fRatioEff := DINT_TO_REAL(nNumEff) / DINT_TO_REAL(nDenEff); // 分母已验非零，防除零
                    ELSE
                        bFaultLatch := TRUE;
                        uErrorId    := 16#0004_0250;         // 【故障级】连续更新传入非法比值
                        eState      := E_DL_GearState.eFault;
                    END_IF
                ELSE
                    uErrorId := 16#0004_0131;                // 【信息级】未开放连续更新时改比值被拒
                END_IF
            END_IF
            // 相位累计（同上，主静止冻结）
            IF ABS(fMasterVel) > DL_GEAR_EPS THEN
                fPhaseErrInt := fPhaseErrInt + (fMasterPosNow - fLastMasterPos) * fRatioEff
                                - (fSlavePosNow - fLastSlavePos);
            ELSE
                uErrorId := 16#0004_0130;                    // 【信息级】主轴静止、相位跟踪冻结
            END_IF
            fCompTerm := 0.0;
            IF (ABS(fPhaseGain) > DL_GEAR_EPS) AND (fPhaseMaxEff > DL_GEAR_EPS) THEN
                fCompTerm := LIMIT(-fPhaseMaxEff, fPhaseGain * fPhaseErrInt, fPhaseMaxEff);
            END_IF
            fTargetCmd := fMasterVel * fRatioEff + fCompTerm;
            IF (fVelLimitEff > DL_GEAR_EPS) AND (ABS(fTargetCmd) > fVelLimitEff) THEN
                fTargetCmd := LIMIT(-fVelLimitEff, fTargetCmd, fVelLimitEff);
                uErrorId   := 16#0004_0132;                  // 【信息级】限速钳位
            END_IF
            // 已啮合段仍以加速度限斜率跟随，防止比值阶跃造成冲击
            fStepMax := fAccEff * fDtS;
            fCmdRamp := fCmdRamp + LIMIT(-fStepMax, fTargetCmd - fCmdRamp, fStepMax);
            fSlaveSpeedCmd := fCmdRamp;
            IF ABS(fCmdRamp - fLastSentCmd) > DL_GEAR_RESEND_EPS THEN
                IF NOT iSlave.MoveVelocity(fVel := fCmdRamp, fAcc := fAccEff) THEN
                    bFaultLatch := TRUE;
                    uErrorId    := 16#0004_0251;             // 【故障级】从轴速度指令被拒
                    fCmdRamp    := 0.0;
                    fSlaveSpeedCmd := 0.0;
                    eState      := E_DL_GearState.eFault;
                ELSE
                    fLastSentCmd := fCmdRamp;
                END_IF
            END_IF
        END_IF

    E_DL_GearState.eDisengaging:                             // 脱开：按减速度受控降速至零后单发停止
        bBusy   := TRUE;
        bActive := FALSE;
        IF iSlave.bError THEN
            bFaultLatch := TRUE;
            uErrorId    := 16#0004_0252;                     // 【故障级】从轴故障中断耦合
            fCmdRamp    := 0.0;
            fSlaveSpeedCmd := 0.0;
            eState      := E_DL_GearState.eFault;
        ELSE
            fStepMax := fDecEff * fDtS;
            fCmdRamp := fCmdRamp - LIMIT(-fStepMax, fCmdRamp, fStepMax); // 朝零收敛，单拍降幅不超 减速度×周期
            IF ABS(fCmdRamp) <= DL_GEAR_EPS THEN
                fCmdRamp       := 0.0;
                fSlaveSpeedCmd := 0.0;
                iSlave.Stop();                               // 指令归零后发一次停止（本拍唯一一次轴调用，随即退态不复发）
                bBusy       := FALSE;
                eState      := E_DL_GearState.eIdle;
            ELSE
                fSlaveSpeedCmd := fCmdRamp;
                IF ABS(fCmdRamp - fLastSentCmd) > DL_GEAR_RESEND_EPS THEN
                    IF NOT iSlave.MoveVelocity(fVel := fCmdRamp, fAcc := fDecEff) THEN
                        bFaultLatch := TRUE;
                        uErrorId    := 16#0004_0251;         // 【故障级】脱开减速指令被拒
                        fCmdRamp    := 0.0;
                        fSlaveSpeedCmd := 0.0;
                        eState      := E_DL_GearState.eFault;
                    ELSE
                        fLastSentCmd := fCmdRamp;
                    END_IF
                END_IF
            END_IF
        END_IF

    E_DL_GearState.eFault:                                   // 故障锁存：仅复位沿可退出
        bInGear        := FALSE;
        bBusy          := FALSE;
        bActive        := FALSE;
        fCmdRamp       := 0.0;
        fSlaveSpeedCmd := 0.0;
        bStopIssued    := FALSE;
        IF fbTrigReset.Q THEN
            bFaultLatch := FALSE;                            // 唯一解除路径
            uErrorId    := 0;
            eState      := E_DL_GearState.eIdle;
        END_IF

    ELSE                                                     // 非法状态兜底（本块专用码）
        bFaultLatch := TRUE;
        uErrorId    := 16#0004_0299;                         // 【故障级】非法状态兜底
        bInGear     := FALSE;
        bBusy       := FALSE;
        bActive     := FALSE;
        fCmdRamp    := 0.0;
        fSlaveSpeedCmd := 0.0;
        eState      := E_DL_GearState.eFault;

END_CASE

// 段 10｜相位基准推进：无论是否耦合都推进一拍，保证增量口径唯一、重新啮合不产生伪增量
fLastMasterPos := fMasterPosNow;                         // 主轴位置基准推进 [mm]
fLastSlavePos  := fSlavePosNow;                          // 从轴位置基准推进 [mm]

// 段 11｜出口映射（派生式，信息级码不参与 bError）
bError       := (eState = E_DL_GearState.eFault);
bInGear      := (eState = E_DL_GearState.eInGear);
bBusy        := (eState = E_DL_GearState.eSynchronizing) OR (eState = E_DL_GearState.eInGear)
                OR (eState = E_DL_GearState.eDisengaging);
bActive      := (eState = E_DL_GearState.eSynchronizing) OR (eState = E_DL_GearState.eInGear);
fRatio       := fRatioEff;
fPhaseError  := fPhaseErrInt;

END_FUNCTION_BLOCK

(* ---- FB_DL_FlyingShearSync.st ---- *)
(*
    FB_DL_FlyingShearSync —— 飞剪同步控制器（加速进入 → 线速同步跟踪 → 剪切触发 → 减速退出）
    ------------------------------------------------------------------
    组件名称  : FB_DL_FlyingShearSync
    分类      : DL_Motion / Synchronization
    前缀      : FB_DL_
    版本      : 1.0.0
    溯源      : 借鉴点 —— PLCopen 对「飞剪 / 飞锯属同步应用」的公开分类事实，
                以及「同步窗 + 速度匹配」的参数域组织方式。
                本件只借**分类事实与参数域组织**，同步区插补数学 / 状态机 /
                码位 100% clean-room 自有，不自造轴状态枚举（轴状态归运动层，
                R31 家族高危区纪律），不引用任何轴接口。
                clean-room 声明 —— 零代码行复制；定时与沿检测仅用 IEC 61131-3
                标准库 TON / R_TRIG，数学仅用标准运算符与 ABS / MAX。
                许可证 —— 本件 MIT；来源标签 t1-6-plcopen 仅指规范文档公开语义，
                规范文本不属代码，无许可继承关系。
    平台      : 纯 IEC 61131-3，CODESYS 3.5 / TwinCAT 3 / InoProShop / Machine Expert 通用
    作者      : 道莅代码库 · PLC编程专家（R71 构建轮 · 批 2 · 序号 5）
    ------------------------------------------------------------------
    功能说明  : 速度级飞剪四段顺控（本件出口为**刀轴速度指令**，非位置指令）：
                eIdle 待机（刀速 0，等切剪请求上升沿）→ eAccel 斜坡加速
                （以 fAccel 向产品线速 fProductVel 逼近，速度差进入 fSyncTol
                即转同步）→ eSyncTrack 线速同步跟踪（刀速直接跟随线速，刀行
                进积分位置进入同步窗 [fShearLen - fSyncWinLen, fShearLen] 后
                受理切剪）→ eCutFire 剪切触发（单拍脉冲，R24 / R187 口径：
                内部 _bCutPulse 置位 → 段 10 统一出口映射单拍，次拍段 1 清零）
                → eDecel 斜坡退窗（以 fDecel 归零）→ eIdle。
                切剪受理规则（计划口径）：bCutReq 上升沿在 eIdle 启动周期并
                预武装 _bCutArmed；在 eSyncTrack 到达即受理（更新武装）；在
                eAccel / eCutFire / eDecel 到达即拒收并计数（信息级，不排队）。
                窗满未剪：eSyncTrack 中刀行进越过 fShearLen 仍未触发 → 信息级
                跳过、撤销武装、强制进 eDecel 清窗（同拍竞态闸：bCutReq 受理
                与窗满判定在同一 CASE 拍内完成，禁跨拍双判）。
                斜坡积分口径（R38）：每拍增量 = 加 / 减速度 × 扫描周期
                （tCycle 引脚注入，无魔法数），运算基于上一拍锁存副本
                _fKnifeCmd，出口单点映射（R191 名实双出口）。
                超时监控（R40）：单实例 _tonPhase，PT 由当前相逐相选择
                （eAccel → tAccelMax，eSyncTrack → tSyncMax，eDecel →
                tDecelMax，段 8 无条件调用），相切换时 IN 随条件清零复位，
                **不跨相累计**（定时器纪律：单定时器逐相 PT，已声明选型）。
                失能语义（R57 / R303）：bEn = FALSE → 速度指令**单拍安全归零**
                （不走斜坡：本件出口为速度指令，斜坡语义由驱动器自身承担，
                停机相输出清零优先于斜坡，安全侧不延时）、状态回 eIdle、
                剪切输出清零；锁存故障不被失能清除，仅 bReset 上升沿解除。
    错误码    : 16#0002_3790 组态非法（切长 / 窗长非正、切长 < 窗长、加速度 /
                            减速度 / 容差非正、扫描周期 / 超时非正、任一非有限），
                            锁存 —— 故障级
                16#0002_3791 加速相超时（未能匹配线速），锁存 —— 故障级
                16#0002_3792 减速相超时（未能归零），锁存 —— 故障级
                16#0002_3793 非法相枚举（CASE ELSE 兜底），锁存 —— 故障级
                16#0002_3798 同步跟踪相超时（窗积分停滞 / 迟迟未到窗），锁存
                            —— 故障级
                16#0002_3794 同步窗满未触发剪切（窗内无有效受理请求），本次跳过
                            进减速 —— 信息级，不置 bError
                16#0002_3795 切剪请求被拒收（非受理相到达），已计数 —— 信息级，
                            不置 bError
                16#0002_3796 产品线速无效（非有限 / 负值），待机相拒收不启动
                            —— 信息级，不置 bError
                16#0002_3797 周期中产品线速失效（非有限 / 负值），锁存停机
                            —— 故障级
    码位总账  : 3790 / 3791 / 3792 / 3793 / 3797 / 3798 用（均故障级）
                3794 / 3795 / 3796 用（信息级，bError 恒 FALSE）
    状态机    : ENUM E_DL_FssPhase 六态，CASE 全覆盖 + ELSE 兜底（锁存 3793
                回 eFault）。迁移表见功能说明；bReset 上升沿：解锁存 →
                eIdle 并清刀速 / 刀位 / 武装（唯一可到达的解除边，R188）。
    边界与披露: 一 组态判据逐项点名（R272）：fShearLen / fSyncWinLen / fAccel /
                   fDecel / fSyncTol 五个 LREAL 全部纳入非有限闸；fSyncWinLen
                   <= 0、fShearLen <= 0、fShearLen < fSyncWinLen（同步窗长于
                   切长即无加速段可言）拦截；fAccel <= 0 / fDecel <= 0 /
                   fSyncTol <= 0 拦截；tCycle / tAccelMax / tDecelMax 非正拦截；
                二 线速守卫：fProductVel 非有限或 < 0.0，待机相拒收（3796，
                   不启动不发指令）；周期中失效锁存（3797，指令归零安全相）；
                   线速 = 0 合法（产品静止，刀速同步为 0，窗积分停滞，由超时
                   收口，头注释声明该边界行为）；
                三 失能相输出清零（R57）：fKnifeVelCmd / bCutTrig 全清零 +
                   状态回 eIdle；锁存相同样清零（失效 / 故障相回夹执行输出）；
                四 剪切脉冲为单拍（R24 / R187 两段式：CASE 内只写内部
                   _bCutPulse，段 10 统一出口映射，段 1 预清零收尾）；
                五 同拍双窗配比约束（R100）：无内建双窗，tAccelMax / tDecelMax
                   与 tCycle 的配比约束为「超时值 >= 2 × tCycle」，否则超时
                   判据可能在相驻留不足两拍时误触发 —— 由组态闸以
                   tAccelMax < 2 * tCycle 拦截（3790）；
                六 定时器 _tonPhase 与沿实例 _rtCut / _rtReset 均无条件周期调用；
                七 计数器 uCutRejCnt 饱和不回绕（增量前预判，R28-3 口径）；
                八 零全局变量、零 VAR_EXTERNAL、零物理地址、零数组下标。
    分工声明  : FB_DL_FlyingCutSync（R37，DL_Motion 同族最近邻）为**位置取模**
                切窗判据件：消费主轴位置、按切长取模计算相位、窗内判同步
                误差后发下刀脉冲，不带加 / 减速斜坡与速度指令出口；本件为
                **速度指令级**四段顺控件：消费产品线速、输出刀轴速度指令，
                两者入口 / 出口契约不同，互引分工不互代（本件立项时按
                R327 词根邻件扫描补记此边界）。FB_DL_LabelApplySync（贴标
                同步）、FB_DL_RotaryIndexModulo（分度回转）为其余同族邻件。
    修订记录  : 2026-11-22 v1.0.0 首次入库（R71 构建轮 · 批 2 · 序号 5）
*)
TYPE E_DL_FssPhase :
(
    eIdle      := 0,   (* 待机，刀速 0，等切剪请求上升沿 / idle, knife at zero, waiting for a cut request edge *)
    eAccel     := 10,  (* 斜坡加速相（向产品线速逼近）/ the accel phase, ramping toward the product speed *)
    eSyncTrack := 20,  (* 线速同步跟踪相（速度跟随 + 刀行进积分 + 同步窗判定）/ the sync track phase, speed follow plus travel integration plus window verdict *)
    eCutFire   := 30,  (* 剪切触发相（单拍脉冲，驻留一拍）/ the cut fire phase, a one scan single pulse *)
    eDecel     := 40,  (* 斜坡减速相（退窗归零）/ the decel phase, ramping back to zero *)
    eFault     := 50   (* 故障相（锁存待复位）/ the fault phase, latched for a reset *)
);
END_TYPE

FUNCTION_BLOCK FB_DL_FlyingShearSync
VAR_INPUT
    bEn         : BOOL := TRUE;            (* 使能，[标志]，FALSE 时指令单拍归零并回待机（R57）/ the enable, FALSE zeroes the command at once and returns to idle *)
    bReset      : BOOL := FALSE;           (* 故障复位（上升沿有效），[标志] / the fault reset, rising edge effective *)
    bCutReq     : BOOL := FALSE;           (* 切剪请求（上升沿启动 / 受理），[标志] / the cut request, rising edge starts or is accepted *)
    fProductVel : LREAL := 0.0;            (* 产品线速，[mm/s]，须 >= 0.0，非有限拒收 / the product line speed, must be non negative and finite *)
    fShearLen   : LREAL := 1000.0;         (* 切长（刀行进目标里程），[mm]，须 >= fSyncWinLen / the shear length, the knife travel target *)
    fSyncWinLen : LREAL := 50.0;           (* 同步窗长（切长尾段允许剪切窗口），[mm]，须 > 0 且 <= fShearLen / the sync window length *)
    fAccel      : LREAL := 5000.0;         (* 加速度，[mm/s²]，须 > 0 / the acceleration *)
    fDecel      : LREAL := 5000.0;         (* 减速度，[mm/s²]，须 > 0 / the deceleration *)
    fSyncTol    : LREAL := 5.0;            (* 速度匹配容差，[mm/s]，须 > 0 / the speed match tolerance *)
    tCycle      : TIME := T#10MS;          (* 扫描周期，[ms]，须 > 0（斜坡积分基值）/ the scan cycle, the ramp integration base *)
    tAccelMax   : TIME := T#5S;            (* 加速相超时，[ms]，须 >= 2 * tCycle / the accel phase timeout *)
    tSyncMax    : TIME := T#10S;           (* 同步跟踪相超时，[ms]，须 >= 2 * tCycle（窗积分停滞的收口）/ the sync track phase timeout *)
    tDecelMax   : TIME := T#5S;            (* 减速相超时，[ms]，须 >= 2 * tCycle / the decel phase timeout *)
END_VAR
VAR_OUTPUT
    eState      : E_DL_FssPhase := E_DL_FssPhase.eIdle; (* 相状态出口，[相] / the phase outlet *)
    fKnifeVelCmd: LREAL;                   (* 刀轴速度指令，[mm/s]，恒 >= 0 / the knife axis velocity command, always non negative *)
    bCutTrig    : BOOL;                    (* 剪切触发脉冲（单拍），[标志] / the cut trigger pulse, single scan *)
    uCutRejCnt  : UDINT;                   (* 切剪请求拒收计数（饱和不回绕）/ the rejected cut request counter, saturating *)
    bValid      : BOOL;                    (* 出口可信（非锁存故障相），[标志] / the outlets trustworthy *)
    bError      : BOOL;                    (* 故障标志，锁存故障时为 TRUE / the fault flag, raised while latched *)
    nErrCode    : UDINT;                   (* 错误码，0 = 正常，锁存回放 / the error id, 0 = ok, replayed from the latch *)
END_VAR
VAR
    _rtCut      : R_TRIG;                  (* 切剪请求上升沿实例（无条件调用）/ the cut request rising edge instance *)
    _rtReset    : R_TRIG;                  (* 复位上升沿实例（无条件调用）/ the reset rising edge instance *)
    _tonPhase   : TON;                     (* 相超时计时实例（单定时器逐相 PT，无条件调用）/ the phase timeout timer, per phase PT *)
    _ePhase     : E_DL_FssPhase := E_DL_FssPhase.eIdle; (* 相状态寄存器 / the internal phase register *)
    _bFault     : BOOL;                    (* 故障锁存位，仅 bReset 上升沿解除 / the latched fault bit *)
    _nCodeLatch : UDINT;                   (* 锁存成因码，故障期回放 / the latched cause code, replayed *)
    _bCfgBad    : BOOL;                    (* 组态非法标志（逐拍重算）/ the configuration fault flag *)
    _bVelBad    : BOOL;                    (* 线速无效标志（逐拍重算）/ the velocity fault flag *)
    _bCutArmed  : BOOL;                    (* 切剪武装位（请求已受理待窗内触发）/ the cut armed flag, a request accepted and waiting for the window *)
    _bCutPulse  : BOOL;                    (* 剪切脉冲内部位（段 10 统一映射，R187）/ the internal cut pulse bit *)
    _fKnifeCmd  : LREAL;                   (* 刀速指令锁存副本（上一拍，R38），[mm/s] / the latched knife command copy, the previous scan *)
    _fKnifePos  : LREAL;                   (* 刀行进积分位置（本周期起点起算），[mm] / the integrated knife travel position *)
    _fDtSec     : LREAL;                   (* 扫描周期秒值（斜坡基值），[s] / the scan cycle in seconds *)
    _fAccStep   : LREAL;                   (* 每拍加速度增量，[mm/s] / the per scan acceleration increment *)
    _fDecStep   : LREAL;                   (* 每拍减速度增量，[mm/s] / the per scan deceleration increment *)
    _bInWin     : BOOL;                    (* 刀位在同步窗内标志，[标志] / the knife sits inside the sync window *)
    _tPhasePt   : TIME;                    (* 相计时器 PT 当前值（逐相选择）/ the timer PT for the current phase *)
    _bTimerIn   : BOOL;                    (* 相计时器 IN 条件（显式条件）/ the timer IN condition *)
END_VAR
VAR CONSTANT
    DL_FSS_FMAX : LREAL := 1.0E30;         (* 非有限筛查幅值上限，[mm 或 mm/s 或 mm/s²] / the finiteness screening cap *)
    DL_FSS_CMAX : UDINT := 16#FFFF_FFFE;   (* 拒收计数饱和上限（增量前预判）/ the reject counter saturation cap, pre-increment check *)
END_VAR

// 段 1｜出口预置（R256 统一出口预置 + 单拍位两段式的第一段）/ segment 1, preset every outlet
eState       := _ePhase;                   // 相出口先镜像寄存器 / mirror the phase register first
bCutTrig     := FALSE;                     // 剪切脉冲预清零（单拍收尾）/ preset the cut pulse false, single scan tail
bValid       := TRUE;                      // 可用标志预置真（故障相再清）/ preset valid true, cleared in the fault phase
bError       := FALSE;                     // 故障标志预清零 / preset the error flag false
nErrCode     := 0;                         // 错误码预置无错 / preset the code to zero
_bCutPulse   := FALSE;                     // 内部脉冲位预清零（次拍清，R187①）/ preset the internal pulse false, cleared next scan
_bTimerIn    := FALSE;                     // 计时条件预清零 / preset the timer condition false
_tPhasePt    := tAccelMax;                 // 计时 PT 预置缺省值 / preset the timer PT to the default

// 段 2｜沿检测实例无条件调用（规则 ⑦）/ segment 2, the edge instances, called unconditionally
_rtCut(CLK := bCutReq);                    // 切剪请求沿，每周期无条件刷新 / the cut request edge, refreshed every scan
_rtReset(CLK := bReset);                   // 复位沿，每周期无条件刷新 / the reset edge, refreshed every scan

// 段 3｜复位解除：唯一可到达的锁存解除边（R188）/ segment 3, the only latch release edge
IF _rtReset.Q THEN                         // 复位上升沿 / the reset rising edge
    _bFault     := FALSE;                  // 解除故障锁存 / release the fault latch
    _nCodeLatch := 0;                      // 清锁存码 / clear the latched code
    _ePhase     := E_DL_FssPhase.eIdle;    // 回待机相（安全相）/ back to the safe idle phase
    _fKnifeCmd  := 0.0;                    // 刀速指令归零 / zero the knife command
    _fKnifePos  := 0.0;                    // 刀行进积分清零 / clear the travel integration
    _bCutArmed  := FALSE;                  // 撤销切剪武装 / disarm the cut request
    _bInWin     := FALSE;                  // 清窗标志 / clear the window flag
END_IF

// 段 4｜组态守卫（边界一逐项点名 + 配比约束边界五，R272）/ segment 4, the configuration guard
_bCfgBad := (fShearLen <= 0.0)                                           // 切长非正 / a non positive shear length
         OR (fSyncWinLen <= 0.0)                                         // 同步窗长非正 / a non positive window length
         OR (fShearLen < fSyncWinLen)                                    // 切长小于窗长（无加速段可言）/ the shear length under the window length
         OR (fAccel <= 0.0)                                              // 加速度非正 / a non positive acceleration
         OR (fDecel <= 0.0)                                              // 减速度非正 / a non positive deceleration
         OR (fSyncTol <= 0.0)                                            // 匹配容差非正 / a non positive tolerance
         OR (tAccelMax < (tCycle + tCycle))                              // 加速超时小于两倍扫描周期（配比约束）/ the accel timeout under two scans
         OR (tSyncMax < (tCycle + tCycle))                               // 同步超时小于两倍扫描周期 / the sync timeout under two scans
         OR (tDecelMax < (tCycle + tCycle))                              // 减速超时小于两倍扫描周期 / the decel timeout under two scans
         OR (fShearLen <> fShearLen) OR ((fShearLen - fShearLen) <> 0.0) OR (ABS(fShearLen) > DL_FSS_FMAX)
         OR (fSyncWinLen <> fSyncWinLen) OR ((fSyncWinLen - fSyncWinLen) <> 0.0) OR (ABS(fSyncWinLen) > DL_FSS_FMAX)
         OR (fAccel <> fAccel) OR ((fAccel - fAccel) <> 0.0) OR (ABS(fAccel) > DL_FSS_FMAX)
         OR (fDecel <> fDecel) OR ((fDecel - fDecel) <> 0.0) OR (ABS(fDecel) > DL_FSS_FMAX)
         OR (fSyncTol <> fSyncTol) OR ((fSyncTol - fSyncTol) <> 0.0) OR (ABS(fSyncTol) > DL_FSS_FMAX);

// 段 5｜线速守卫：非有限或负值即无效（待机拒收 / 周期中锁存，边界二）/ segment 5, the velocity guard
_bVelBad := (fProductVel <> fProductVel) OR ((fProductVel - fProductVel) <> 0.0) // 线速非有限 / the speed non finite
         OR (fProductVel < 0.0)                                  // 线速为负 / a negative speed
         OR (ABS(fProductVel) > DL_FSS_FMAX);                    // 线速超幅值筛查 / the speed over the screening cap

// 段 6｜首次成因锁存（故障期不重推断，回放锁存码，R189）/ segment 6, the first-cause latch
IF NOT _bFault THEN                        // 未锁存才登记成因 / a cause is registered only while not latched
    IF _bCfgBad THEN                       // 组态非法优先归因（根因）/ the configuration first, the root cause
        _bFault     := TRUE;               // 置锁存 / latch it
        _nCodeLatch := 16#0002_3790;       // 故障级：组态非法 / fault level: an illegal configuration
        _ePhase     := E_DL_FssPhase.eFault; // 迁入故障相 / enter the fault phase
    ELSIF _bVelBad AND (_ePhase <> E_DL_FssPhase.eIdle) THEN // 周期中线速失效 / the speed failed mid cycle
        _bFault     := TRUE;               // 置锁存 / latch it
        _nCodeLatch := 16#0002_3797;       // 故障级：线速失效停机 / fault level: the speed failed in cycle
        _ePhase     := E_DL_FssPhase.eFault; // 迁入故障相 / enter the fault phase
    END_IF
END_IF

// 段 7｜斜坡基值换算（TIME 显式转 ms 再转秒，不依赖平台 TIME_TO_LREAL 语义差）/ segment 7, the ramp base conversion
_fDtSec   := DINT_TO_LREAL(TIME_TO_DINT(tCycle)) / 1000.0; // 扫描周期秒值（除子为常量 1000.0，无除零面）/ the cycle in seconds, a constant divisor
_fAccStep := fAccel * _fDtSec;             // 每拍加速增量，[mm/s] / the per scan accel increment
_fDecStep := fDecel * _fDtSec;             // 每拍减速增量，[mm/s] / the per scan decel increment

// 段 8｜相计时器 PT 选择与无条件调用（规则 ⑦，选相不依赖可跳过分支）/ segment 8, the timer PT selection and the unconditional call
IF _ePhase = E_DL_FssPhase.eAccel THEN     // 加速相 / the accel phase
    _tPhasePt := tAccelMax;                // 加速超时值 / the accel timeout
    _bTimerIn := TRUE;                     // 相内计时有效 / the timer runs inside the phase
ELSIF _ePhase = E_DL_FssPhase.eSyncTrack THEN // 同步跟踪相 / the sync track phase
    _tPhasePt := tSyncMax;                 // 同步超时值（窗积分停滞收口）/ the sync timeout
    _bTimerIn := TRUE;                     // 相内计时有效 / the timer runs
ELSIF _ePhase = E_DL_FssPhase.eDecel THEN  // 减速相 / the decel phase
    _tPhasePt := tDecelMax;                // 减速超时值 / the decel timeout
    _bTimerIn := TRUE;                     // 相内计时有效 / the timer runs
ELSE                                       // 其余相不参与计时（缺省分支，非状态机 ELSE）/ the other phases do not time
    _tPhasePt := tAccelMax;                // 缺省 PT，保证 PT 恒有定义 / a default PT, always defined
    _bTimerIn := FALSE;                    // 计时条件清零 / the timer condition cleared
END_IF
_tonPhase(IN := _bTimerIn, PT := _tPhasePt); // 每周期无条件调用 / called every scan without exception

// 段 8b｜失能与故障相输出回夹（R57 停机相输出清零，先于状态机执行）/ segment 8b, the disable and fault output clamping
IF _bFault THEN                            // 锁存故障相 / the latched fault phase
    _fKnifeCmd := 0.0;                     // 刀速指令归零（回夹执行输出）/ zero the command, clamp the outlet
    _bCutArmed := FALSE;                   // 撤销武装 / disarm
    _bInWin    := FALSE;                   // 清窗 / clear the window
ELSIF NOT bEn THEN                         // 失能相（操作态，不发码）/ the disabled phase, an operator state
    _fKnifeCmd := 0.0;                     // 失能单拍安全归零（边界三，不走斜坡）/ zeroed at once, no ramp
    _ePhase    := E_DL_FssPhase.eIdle;     // 状态回待机 / back to idle
    _bCutArmed := FALSE;                   // 撤销武装 / disarm
    _bInWin    := FALSE;                   // 清窗 / clear the window
END_IF

// 段 9｜相状态机（ENUM + CASE + ELSE 兜底，仅运行许可时执行）/ segment 9, the phase machine, run permit only
IF bEn AND NOT _bFault THEN                // 运行许可成立 / the run permit holds
CASE _ePhase OF
    E_DL_FssPhase.eIdle:                   // 待机相 / the idle phase
        IF _bVelBad THEN                   // 线速无效（待机拒收，不发指令）/ the speed invalid, refused at idle
            nErrCode := 16#0002_3796;      // 信息级：待机拒收（不置 bError，R45）/ info level: refused at idle
        ELSIF _rtCut.Q THEN                // 切剪请求上升沿（启动周期并武装）/ a cut request edge starts the cycle
            _bCutArmed := TRUE;           // 预武装本请求 / arm this request
            _fKnifePos := 0.0;            // 刀行进积分清零（周期起点）/ clear the travel integration
            _ePhase    := E_DL_FssPhase.eAccel; // 进入加速相 / enter the accel phase
        END_IF
    E_DL_FssPhase.eAccel:                  // 加速相 / the accel phase
        IF _rtCut.Q THEN                   // 非受理相请求到达 → 拒收计数 / a request in a non accepting phase, refused
            IF uCutRejCnt < DL_FSS_CMAX THEN // 饱和不回绕（增量前预判）/ saturating, no wrap
                uCutRejCnt := uCutRejCnt + 1; // 拒收计数递增 / increment the reject counter
            END_IF
            nErrCode := 16#0002_3795;      // 信息级：请求被拒收 / info level: the request refused
        END_IF
        IF ABS(_fKnifeCmd - fProductVel) <= fSyncTol THEN // 速度差进入容差带 / the speed gap inside the tolerance
            _fKnifeCmd := fProductVel;     // 贴合线速（消除残余差）/ snap onto the line speed
            _ePhase    := E_DL_FssPhase.eSyncTrack; // 进入同步跟踪相 / enter the sync track phase
        ELSE                               // 尚未匹配 / not matched yet
            _fKnifeCmd := _fKnifeCmd + _fAccStep; // 斜坡上抬（基于上一拍副本，R38）/ ramp up from the latched copy
            IF _fKnifeCmd > fProductVel THEN   // 越过目标（超调钳位，贴线速后不再上抬）/ over the target, clamp the overshoot
                _fKnifeCmd := fProductVel;     // 钳到目标 / clamp to the target
            END_IF
        END_IF
        _fKnifePos := _fKnifePos + _fKnifeCmd * _fDtSec; // 刀行进积分（加速段亦前进）/ the travel integration, the knife advances
        IF _tonPhase.Q THEN                // 加速相超时（归因唯一 3791）/ the accel phase timed out
            _bFault     := TRUE;           // 锁存故障 / latch the fault
            _nCodeLatch := 16#0002_3791;   // 故障级：加速超时 / fault level: the accel timed out
            _ePhase     := E_DL_FssPhase.eFault; // 迁入故障相 / enter the fault phase
        END_IF
    E_DL_FssPhase.eSyncTrack:              // 同步跟踪相 / the sync track phase
        _fKnifeCmd := fProductVel;         // 速度直接跟随线速（同步段不再斜坡）/ follow the line speed directly
        _fKnifePos := _fKnifePos + _fKnifeCmd * _fDtSec; // 刀行进积分 / the travel integration
        _bInWin    := (_fKnifePos >= (fShearLen - fSyncWinLen)); // 同步窗判定（闭区间下界）/ the window verdict, a closed lower bound
        IF _rtCut.Q THEN                   // 受理相请求到达 → 更新武装 / a request in the accepting phase, arm it
            _bCutArmed := TRUE;            // 受理 / accepted
        END_IF
        IF _bCutArmed AND _bInWin AND (ABS(_fKnifeCmd - fProductVel) <= fSyncTol) THEN // 窗内 + 已匹配 + 已武装 → 触发
            _ePhase := E_DL_FssPhase.eCutFire; // 进入剪切触发相（下拍发脉冲）/ enter the cut fire phase
        ELSIF _fKnifePos >= fShearLen THEN // 窗满未剪（同拍竞态闸：本拍事件已先消化）/ the window passed without a cut
            _bCutArmed := FALSE;           // 撤销武装 / disarm
            nErrCode   := 16#0002_3794;    // 信息级：窗满跳过 / info level: skipped
            _ePhase    := E_DL_FssPhase.eDecel; // 强制进减速清窗 / force the decel phase to clear the window
        ELSIF _tonPhase.Q THEN             // 同步跟踪相超时（归因唯一 3798，窗积分停滞的收口）/ the sync track timed out
            _bFault     := TRUE;           // 锁存故障 / latch the fault
            _nCodeLatch := 16#0002_3798;   // 故障级：同步超时 / fault level: the sync track timed out
            _ePhase     := E_DL_FssPhase.eFault; // 迁入故障相 / enter the fault phase
        END_IF
    E_DL_FssPhase.eCutFire:                // 剪切触发相（驻留一拍）/ the cut fire phase, one scan
        _bCutPulse := TRUE;                // 内部脉冲置位（段 10 统一映射，R187）/ set the internal pulse, mapped at segment 10
        _ePhase    := E_DL_FssPhase.eDecel; // 次拍转入减速相 / move to the decel phase next scan
    E_DL_FssPhase.eDecel:                  // 减速相 / the decel phase
        IF _rtCut.Q THEN                   // 非受理相请求到达 → 拒收计数 / a request in a non accepting phase, refused
            IF uCutRejCnt < DL_FSS_CMAX THEN // 饱和不回绕 / saturating
                uCutRejCnt := uCutRejCnt + 1; // 拒收计数递增 / increment the counter
            END_IF
            nErrCode := 16#0002_3795;      // 信息级：请求被拒收 / info level: refused
        END_IF
        _fKnifeCmd := _fKnifeCmd - _fDecStep; // 斜坡下降（基于上一拍副本，R38）/ ramp down from the latched copy
        IF _fKnifeCmd <= 0.0 THEN          // 已归零（MAX 钳位结果，非浮点判等）/ zeroed via the MAX clamp, no float equality
            _fKnifeCmd := 0.0;          // 精确归零 / exact zero
            _fKnifePos := 0.0;           // 刀位清零（下周期起点复位）/ clear the travel position
            _bInWin    := FALSE;         // 清窗 / clear the window
            _ePhase    := E_DL_FssPhase.eIdle; // 回待机 / back to idle
        END_IF
        IF _tonPhase.Q THEN                // 减速相超时（归因唯一 3792）/ the decel phase timed out
            _bFault     := TRUE;           // 锁存故障 / latch the fault
            _nCodeLatch := 16#0002_3792;   // 故障级：减速超时 / fault level: the decel timed out
            _ePhase     := E_DL_FssPhase.eFault; // 迁入故障相 / enter the fault phase
        END_IF
    E_DL_FssPhase.eFault:                  // 故障相（锁存保持，输出回夹已在段 8b 执行）/ the fault phase, outlets clamped at 8b
        bValid   := FALSE;                 // 出口不可信 / the outlets not trustworthy
        bError   := TRUE;                  // 故障标志置位 / raise the fault flag
        nErrCode := _nCodeLatch;           // 回放锁存码（不按当下输入重推断）/ replay the latched code
    ELSE                                   // 非法枚举兜底（回安全相 + 置码，规则 ⑥）/ the illegal enumeration guard
        _bFault     := TRUE;               // 置锁存 / latch it
        _nCodeLatch := 16#0002_3793;       // 故障级：非法相枚举 / fault level: an illegal phase value
        _ePhase     := E_DL_FssPhase.eFault; // 回安全相（故障相）/ force the safe fault phase
        bValid      := FALSE;              // 出口不可信 / not trustworthy
        bError      := TRUE;               // 故障标志置位（禁静默）/ raise the flag
        nErrCode    := _nCodeLatch;        // 回放锁存码 / replay the latched code
END_CASE
END_IF

// 段 10｜出口映射（名实双出口同源，单点写入，R191）/ segment 10, the outlet mapping
fKnifeVelCmd := _fKnifeCmd;                // 刀速指令出口 = 锁存副本（单点写入）/ the command outlet mirrors the register
bCutTrig     := _bCutPulse AND bEn AND NOT _bFault; // 剪切脉冲单拍出口（失能 / 故障禁发）/ the single scan pulse, gated
eState       := _ePhase;                   // 相出口 = 寄存器（段 9 之后不再触碰）/ the phase outlet, not touched after segment 9
IF _bFault THEN                            // 锁存故障相出口补充（含故障入口拍，指令即时归零回夹）/ the latched fault supplement, including the entry scan
    fKnifeVelCmd := 0.0;                   // 刀速指令归零（回夹执行输出）/ zero the command outlet
    bValid   := FALSE;                     // 出口不可信 / not trustworthy
    bError   := TRUE;                      // 故障标志 / the fault flag
    nErrCode := _nCodeLatch;               // 回放锁存码 / replay the latched code
END_IF
END_FUNCTION_BLOCK
